  movel([0.147187, -1.292502, -2.622642, -0.797245, 1.570796, 1.717984],accel_mss,speed_ms,0,blend_radius_m)
  movel([0.147550, -1.292939, -2.622384, -0.797065, 1.570796, 1.718347],accel_mss,speed_ms,0,blend_radius_m)
  movel([0.147774, -1.294240, -2.621617, -0.796531, 1.570796, 1.718570],accel_mss,speed_ms,0,blend_radius_m)
  movel([0.147672, -1.296185, -2.620466, -0.795737, 1.570796, 1.718469],accel_mss,speed_ms,0,blend_radius_m)
  movel([0.147381, -1.298185, -2.619278, -0.794926, 1.570796, 1.718178],accel_mss,speed_ms,0,blend_radius_m)
  movel([0.149143, -1.296279, -2.620411, -0.795699, 1.570796, 1.719939],accel_mss,speed_ms,0,blend_radius_m)
  movel([0.151055, -1.294467, -2.621483, -0.796439, 1.570796, 1.721852],accel_mss,speed_ms,0,blend_radius_m)
  movel([0.153085, -1.292767, -2.622486, -0.797136, 1.570796, 1.723882],accel_mss,speed_ms,0,blend_radius_m)
  movel([0.155193, -1.291198, -2.623408, -0.797783, 1.570796, 1.725989],accel_mss,speed_ms,0,blend_radius_m)
  movel([0.159402, -1.288061, -2.625242, -0.799086, 1.570796, 1.730199],accel_mss,speed_ms,0,blend_radius_m)
  movel([0.160619, -1.287255, -2.625711, -0.799423, 1.570796, 1.731416],accel_mss,speed_ms,0,blend_radius_m)
  movel([0.161780, -1.286599, -2.626092, -0.799698, 1.570796, 1.732576],accel_mss,speed_ms,0,blend_radius_m)
  movel([0.162826, -1.286172, -2.626340, -0.799877, 1.570796, 1.733623],accel_mss,speed_ms,0,blend_radius_m)
  movel([0.163696, -1.286049, -2.626411, -0.799928, 1.570796, 1.734492],accel_mss,speed_ms,0,blend_radius_m)
  movel([0.164332, -1.286333, -2.626247, -0.799809, 1.570796, 1.735128],accel_mss,speed_ms,0,blend_radius_m)
  movel([0.164662, -1.286984, -2.625868, -0.799536, 1.570796, 1.735459],accel_mss,speed_ms,0,blend_radius_m)
  movel([0.164729, -1.287902, -2.625335, -0.799153, 1.570796, 1.735526],accel_mss,speed_ms,0,blend_radius_m)
  movel([0.164568, -1.288980, -2.624706, -0.798703, 1.570796, 1.735364],accel_mss,speed_ms,0,blend_radius_m)
  movel([0.164219, -1.290117, -2.624041, -0.798231, 1.570796, 1.735015],accel_mss,speed_ms,0,blend_radius_m)
  movel([0.163722, -1.291209, -2.623401, -0.797779, 1.570796, 1.734518],accel_mss,speed_ms,0,blend_radius_m)
  movel([0.163113, -1.292155, -2.622846, -0.797388, 1.570796, 1.733910],accel_mss,speed_ms,0,blend_radius_m)
  movel([0.162431, -1.292853, -2.622435, -0.797101, 1.570796, 1.733227],accel_mss,speed_ms,0,blend_radius_m)
  movel([0.166229, -1.290188, -2.624000, -0.798201, 1.570796, 1.737025],accel_mss,speed_ms,0,blend_radius_m)
  movel([0.168191, -1.288999, -2.624694, -0.798695, 1.570796, 1.738988],accel_mss,speed_ms,0,blend_radius_m)
  movel([0.170182, -1.287929, -2.625319, -0.799141, 1.570796, 1.740979],accel_mss,speed_ms,0,blend_radius_m)
  movel([0.172188, -1.286991, -2.625865, -0.799534, 1.570796, 1.742984],accel_mss,speed_ms,0,blend_radius_m)
  movel([0.174199, -1.286202, -2.626323, -0.799864, 1.570796, 1.744995],accel_mss,speed_ms,0,blend_radius_m)
  movel([0.176204, -1.285580, -2.626683, -0.800126, 1.570796, 1.747000],accel_mss,speed_ms,0,blend_radius_m)
  movel([0.178191, -1.285136, -2.626940, -0.800312, 1.570796, 1.748987],accel_mss,speed_ms,0,blend_radius_m)
  movel([0.179463, -1.285131, -2.626943, -0.800314, 1.570796, 1.750259],accel_mss,speed_ms,0,blend_radius_m)
  movel([0.180721, -1.285520, -2.626718, -0.800151, 1.570796, 1.751518],accel_mss,speed_ms,0,blend_radius_m)
  movel([0.181223, -1.285864, -2.626519, -0.800006, 1.570796, 1.752019],accel_mss,speed_ms,0,blend_radius_m)
  movel([0.181576, -1.286307, -2.626262, -0.799820, 1.570796, 1.752372],accel_mss,speed_ms,0,blend_radius_m)
  movel([0.181734, -1.286851, -2.625946, -0.799592, 1.570796, 1.752530],accel_mss,speed_ms,0,blend_radius_m)
  movel([0.181645, -1.287496, -2.625571, -0.799322, 1.570796, 1.752441],accel_mss,speed_ms,0,blend_radius_m)
  movel([0.181300, -1.288146, -2.625192, -0.799051, 1.570796, 1.752096],accel_mss,speed_ms,0,blend_radius_m)
  movel([0.180775, -1.288760, -2.624834, -0.798795, 1.570796, 1.751571],accel_mss,speed_ms,0,blend_radius_m)
  movel([0.179372, -1.289953, -2.624137, -0.798299, 1.570796, 1.750168],accel_mss,speed_ms,0,blend_radius_m)
  movel([0.177819, -1.290875, -2.623597, -0.797917, 1.570796, 1.748615],accel_mss,speed_ms,0,blend_radius_m)
  movel([0.176195, -1.291571, -2.623189, -0.797629, 1.570796, 1.746991],accel_mss,speed_ms,0,blend_radius_m)
  movel([0.174578, -1.292087, -2.622886, -0.797416, 1.570796, 1.745374],accel_mss,speed_ms,0,blend_radius_m)
  movel([0.176378, -1.292531, -2.622625, -0.797233, 1.570796, 1.747174],accel_mss,speed_ms,0,blend_radius_m)
  movel([0.178306, -1.292768, -2.622485, -0.797136, 1.570796, 1.749103],accel_mss,speed_ms,0,blend_radius_m)
  movel([0.180340, -1.292800, -2.622467, -0.797123, 1.570796, 1.751137],accel_mss,speed_ms,0,blend_radius_m)
  movel([0.182461, -1.292627, -2.622568, -0.797194, 1.570796, 1.753257],accel_mss,speed_ms,0,blend_radius_m)
  movel([0.184182, -1.292297, -2.622762, -0.797330, 1.570796, 1.754979],accel_mss,speed_ms,0,blend_radius_m)
  movel([0.187621, -1.291362, -2.623311, -0.797715, 1.570796, 1.758417],accel_mss,speed_ms,0,blend_radius_m)
  movel([0.189347, -1.291019, -2.623513, -0.797857, 1.570796, 1.760143],accel_mss,speed_ms,0,blend_radius_m)
  movel([0.191271, -1.290783, -2.623651, -0.797955, 1.570796, 1.762067],accel_mss,speed_ms,0,blend_radius_m)
  movel([0.194455, -1.290577, -2.623772, -0.798040, 1.570796, 1.765251],accel_mss,speed_ms,0,blend_radius_m)
  movel([0.195937, -1.290628, -2.623742, -0.798019, 1.570796, 1.766733],accel_mss,speed_ms,0,blend_radius_m)
  movel([0.197036, -1.290857, -2.623608, -0.797924, 1.570796, 1.767833],accel_mss,speed_ms,0,blend_radius_m)
  movel([0.197371, -1.291056, -2.623491, -0.797842, 1.570796, 1.768167],accel_mss,speed_ms,0,blend_radius_m)
  movel([0.197521, -1.291320, -2.623336, -0.797733, 1.570796, 1.768317],accel_mss,speed_ms,0,blend_radius_m)
  movel([0.197462, -1.291654, -2.623140, -0.797595, 1.570796, 1.768258],accel_mss,speed_ms,0,blend_radius_m)
  movel([0.197162, -1.292065, -2.622898, -0.797425, 1.570796, 1.767958],accel_mss,speed_ms,0,blend_radius_m)
  movel([0.196189, -1.292919, -2.622396, -0.797073, 1.570796, 1.766986],accel_mss,speed_ms,0,blend_radius_m)
  movel([0.195007, -1.293687, -2.621944, -0.796758, 1.570796, 1.765803],accel_mss,speed_ms,0,blend_radius_m)
  movel([0.193677, -1.294378, -2.621536, -0.796475, 1.570796, 1.764473],accel_mss,speed_ms,0,blend_radius_m)
  movel([0.192268, -1.294993, -2.621172, -0.796224, 1.570796, 1.763065],accel_mss,speed_ms,0,blend_radius_m)
  movel([0.189469, -1.296012, -2.620569, -0.795808, 1.570796, 1.760265],accel_mss,speed_ms,0,blend_radius_m)
  movel([0.187130, -1.296774, -2.620117, -0.795498, 1.570796, 1.757926],accel_mss,speed_ms,0,blend_radius_m)
  movel([0.188093, -1.297277, -2.619818, -0.795294, 1.570796, 1.758889],accel_mss,speed_ms,0,blend_radius_m)
  movel([0.189142, -1.297667, -2.619586, -0.795136, 1.570796, 1.759938],accel_mss,speed_ms,0,blend_radius_m)
  movel([0.191445, -1.298162, -2.619291, -0.794935, 1.570796, 1.762241],accel_mss,speed_ms,0,blend_radius_m)
  movel([0.193943, -1.298359, -2.619175, -0.794856, 1.570796, 1.764739],accel_mss,speed_ms,0,blend_radius_m)
  movel([0.196543, -1.298358, -2.619175, -0.794856, 1.570796, 1.767339],accel_mss,speed_ms,0,blend_radius_m)
  movel([0.198733, -1.298215, -2.619260, -0.794914, 1.570796, 1.769529],accel_mss,speed_ms,0,blend_radius_m)
  movel([0.205405, -1.297512, -2.619678, -0.795198, 1.570796, 1.776202],accel_mss,speed_ms,0,blend_radius_m)
  movel([0.206582, -1.297609, -2.619621, -0.795159, 1.570796, 1.777379],accel_mss,speed_ms,0,blend_radius_m)
  movel([0.207429, -1.297998, -2.619389, -0.795002, 1.570796, 1.778225],accel_mss,speed_ms,0,blend_radius_m)
  movel([0.207554, -1.298296, -2.619212, -0.794881, 1.570796, 1.778350],accel_mss,speed_ms,0,blend_radius_m)
  movel([0.207384, -1.298662, -2.618994, -0.794733, 1.570796, 1.778180],accel_mss,speed_ms,0,blend_radius_m)
  movel([0.206850, -1.299092, -2.618737, -0.794560, 1.570796, 1.777646],accel_mss,speed_ms,0,blend_radius_m)
  movel([0.205881, -1.299582, -2.618444, -0.794362, 1.570796, 1.776677],accel_mss,speed_ms,0,blend_radius_m)
  movel([0.204309, -1.300170, -2.618093, -0.794126, 1.570796, 1.775105],accel_mss,speed_ms,0,blend_radius_m)
  movel([0.202535, -1.300655, -2.617803, -0.793931, 1.570796, 1.773331],accel_mss,speed_ms,0,blend_radius_m)
  movel([0.200836, -1.300909, -2.617651, -0.793829, 1.570796, 1.771632],accel_mss,speed_ms,0,blend_radius_m)
  movel([0.200100, -1.300910, -2.617650, -0.793829, 1.570796, 1.770896],accel_mss,speed_ms,0,blend_radius_m)
  movel([0.199490, -1.300801, -2.617716, -0.793873, 1.570796, 1.770286],accel_mss,speed_ms,0,blend_radius_m)
  movel([0.201611, -1.302312, -2.616809, -0.793268, 1.570796, 1.772407],accel_mss,speed_ms,0,blend_radius_m)
  movel([0.203973, -1.303547, -2.616066, -0.792776, 1.570796, 1.774769],accel_mss,speed_ms,0,blend_radius_m)
  movel([0.206525, -1.304557, -2.615457, -0.792375, 1.570796, 1.777321],accel_mss,speed_ms,0,blend_radius_m)
  movel([0.209220, -1.305396, -2.614950, -0.792043, 1.570796, 1.780016],accel_mss,speed_ms,0,blend_radius_m)
  movel([0.214839, -1.306755, -2.614126, -0.791507, 1.570796, 1.785635],accel_mss,speed_ms,0,blend_radius_m)
  movel([0.220430, -1.308023, -2.613356, -0.791010, 1.570796, 1.791226],accel_mss,speed_ms,0,blend_radius_m)
  movel([0.221316, -1.308412, -2.613120, -0.790858, 1.570796, 1.792112],accel_mss,speed_ms,0,blend_radius_m)
  movel([0.221557, -1.308760, -2.612908, -0.790722, 1.570796, 1.792354],accel_mss,speed_ms,0,blend_radius_m)
  movel([0.221539, -1.309244, -2.612612, -0.790532, 1.570796, 1.792335],accel_mss,speed_ms,0,blend_radius_m)
  movel([0.221247, -1.309765, -2.612295, -0.790329, 1.570796, 1.792044],accel_mss,speed_ms,0,blend_radius_m)
  movel([0.220033, -1.310912, -2.611593, -0.789884, 1.570796, 1.790829],accel_mss,speed_ms,0,blend_radius_m)
  movel([0.219216, -1.311486, -2.611242, -0.789661, 1.570796, 1.790013],accel_mss,speed_ms,0,blend_radius_m)
  movel([0.217461, -1.312385, -2.610691, -0.789314, 1.570796, 1.788257],accel_mss,speed_ms,0,blend_radius_m)
  movel([0.215610, -1.312982, -2.610324, -0.789083, 1.570796, 1.786407],accel_mss,speed_ms,0,blend_radius_m)
  movel([0.213729, -1.313322, -2.610115, -0.788953, 1.570796, 1.784525],accel_mss,speed_ms,0,blend_radius_m)
  movel([0.211888, -1.313440, -2.610042, -0.788907, 1.570796, 1.782685],accel_mss,speed_ms,0,blend_radius_m)
  movel([0.210157, -1.313379, -2.610079, -0.788930, 1.570796, 1.780953],accel_mss,speed_ms,0,blend_radius_m)
  movel([0.208604, -1.313175, -2.610205, -0.789009, 1.570796, 1.779400],accel_mss,speed_ms,0,blend_radius_m)
  movel([0.207302, -1.312863, -2.610397, -0.789129, 1.570796, 1.778098],accel_mss,speed_ms,0,blend_radius_m)
  movel([0.207188, -1.313311, -2.610121, -0.788957, 1.570796, 1.777984],accel_mss,speed_ms,0,blend_radius_m)
  movel([0.207346, -1.313680, -2.609894, -0.788815, 1.570796, 1.778142],accel_mss,speed_ms,0,blend_radius_m)
  movel([0.207939, -1.314359, -2.609476, -0.788554, 1.570796, 1.778735],accel_mss,speed_ms,0,blend_radius_m)
  movel([0.208657, -1.314923, -2.609128, -0.788338, 1.570796, 1.779454],accel_mss,speed_ms,0,blend_radius_m)
  movel([0.210309, -1.315835, -2.608564, -0.787990, 1.570796, 1.781105],accel_mss,speed_ms,0,blend_radius_m)
  movel([0.213305, -1.317223, -2.607704, -0.787461, 1.570796, 1.784102],accel_mss,speed_ms,0,blend_radius_m)
  movel([0.216384, -1.318478, -2.606925, -0.786986, 1.570796, 1.787181],accel_mss,speed_ms,0,blend_radius_m)
  movel([0.222772, -1.320657, -2.605566, -0.786166, 1.570796, 1.793568],accel_mss,speed_ms,0,blend_radius_m)
  movel([0.224533, -1.321298, -2.605165, -0.785925, 1.570796, 1.795329],accel_mss,speed_ms,0,blend_radius_m)
  movel([0.225622, -1.321824, -2.604836, -0.785729, 1.570796, 1.796418],accel_mss,speed_ms,0,blend_radius_m)
  movel([0.226633, -1.322477, -2.604427, -0.785485, 1.570796, 1.797429],accel_mss,speed_ms,0,blend_radius_m)
  movel([0.227396, -1.323251, -2.603940, -0.785197, 1.570796, 1.798192],accel_mss,speed_ms,0,blend_radius_m)
  movel([0.227749, -1.324134, -2.603385, -0.784870, 1.570796, 1.798546],accel_mss,speed_ms,0,blend_radius_m)
  movel([0.227725, -1.324612, -2.603084, -0.784693, 1.570796, 1.798521],accel_mss,speed_ms,0,blend_radius_m)
  movel([0.227538, -1.325115, -2.602767, -0.784507, 1.570796, 1.798334],accel_mss,speed_ms,0,blend_radius_m)
  movel([0.227164, -1.325643, -2.602434, -0.784312, 1.570796, 1.797961],accel_mss,speed_ms,0,blend_radius_m)
  movel([0.226591, -1.326191, -2.602087, -0.784110, 1.570796, 1.797387],accel_mss,speed_ms,0,blend_radius_m)
  movel([0.225837, -1.326540, -2.601867, -0.783982, 1.570796, 1.796634],accel_mss,speed_ms,0,blend_radius_m)
  movel([0.224871, -1.326699, -2.601766, -0.783924, 1.570796, 1.795668],accel_mss,speed_ms,0,blend_radius_m)
  movel([0.219802, -1.326944, -2.601611, -0.783834, 1.570796, 1.790598],accel_mss,speed_ms,0,blend_radius_m)
  movel([0.218145, -1.326787, -2.601710, -0.783892, 1.570796, 1.788941],accel_mss,speed_ms,0,blend_radius_m)
  movel([0.217459, -1.326589, -2.601836, -0.783964, 1.570796, 1.788255],accel_mss,speed_ms,0,blend_radius_m)
  movel([0.216923, -1.326283, -2.602029, -0.784077, 1.570796, 1.787719],accel_mss,speed_ms,0,blend_radius_m)
  movel([0.218941, -1.328596, -2.600563, -0.783230, 1.570796, 1.789737],accel_mss,speed_ms,0,blend_radius_m)
  movel([0.221308, -1.330580, -2.599299, -0.782510, 1.570796, 1.792105],accel_mss,speed_ms,0,blend_radius_m)
  movel([0.223948, -1.332287, -2.598208, -0.781894, 1.570796, 1.794744],accel_mss,speed_ms,0,blend_radius_m)
  movel([0.226784, -1.333763, -2.597261, -0.781365, 1.570796, 1.797581],accel_mss,speed_ms,0,blend_radius_m)
  movel([0.229318, -1.334606, -2.596719, -0.781064, 1.570796, 1.800115],accel_mss,speed_ms,0,blend_radius_m)
  movel([0.232932, -1.335887, -2.595893, -0.780608, 1.570796, 1.803728],accel_mss,speed_ms,0,blend_radius_m)
  movel([0.234525, -1.336695, -2.595372, -0.780322, 1.570796, 1.805322],accel_mss,speed_ms,0,blend_radius_m)
  movel([0.235653, -1.337610, -2.594780, -0.780000, 1.570796, 1.806450],accel_mss,speed_ms,0,blend_radius_m)
  movel([0.235966, -1.338106, -2.594458, -0.779825, 1.570796, 1.806763],accel_mss,speed_ms,0,blend_radius_m)
  movel([0.236070, -1.338627, -2.594120, -0.779642, 1.570796, 1.806867],accel_mss,speed_ms,0,blend_radius_m)
  movel([0.235936, -1.339175, -2.593764, -0.779450, 1.570796, 1.806733],accel_mss,speed_ms,0,blend_radius_m)
  movel([0.235538, -1.339746, -2.593393, -0.779250, 1.570796, 1.806335],accel_mss,speed_ms,0,blend_radius_m)
  movel([0.234996, -1.340245, -2.593068, -0.779076, 1.570796, 1.805793],accel_mss,speed_ms,0,blend_radius_m)
  movel([0.234397, -1.340669, -2.592792, -0.778928, 1.570796, 1.805193],accel_mss,speed_ms,0,blend_radius_m)
  movel([0.233113, -1.341353, -2.592346, -0.778690, 1.570796, 1.803910],accel_mss,speed_ms,0,blend_radius_m)
  movel([0.231720, -1.341950, -2.591956, -0.778483, 1.570796, 1.802517],accel_mss,speed_ms,0,blend_radius_m)
  movel([0.228948, -1.342826, -2.591382, -0.778180, 1.570796, 1.799744],accel_mss,speed_ms,0,blend_radius_m)
  movel([0.227584, -1.343104, -2.591201, -0.778085, 1.570796, 1.798381],accel_mss,speed_ms,0,blend_radius_m)
  movel([0.229786, -1.344148, -2.590516, -0.777725, 1.570796, 1.800582],accel_mss,speed_ms,0,blend_radius_m)
  movel([0.232093, -1.345031, -2.589935, -0.777422, 1.570796, 1.802889],accel_mss,speed_ms,0,blend_radius_m)
  movel([0.234492, -1.345775, -2.589446, -0.777168, 1.570796, 1.805289],accel_mss,speed_ms,0,blend_radius_m)
  movel([0.236975, -1.346392, -2.589039, -0.776958, 1.570796, 1.807771],accel_mss,speed_ms,0,blend_radius_m)
  movel([0.242140, -1.347324, -2.588424, -0.776642, 1.570796, 1.812936],accel_mss,speed_ms,0,blend_radius_m)
  movel([0.247502, -1.347956, -2.588005, -0.776427, 1.570796, 1.818298],accel_mss,speed_ms,0,blend_radius_m)
  movel([0.248879, -1.348279, -2.587792, -0.776318, 1.570796, 1.819675],accel_mss,speed_ms,0,blend_radius_m)
  movel([0.249326, -1.348656, -2.587542, -0.776191, 1.570796, 1.820123],accel_mss,speed_ms,0,blend_radius_m)
  movel([0.249438, -1.349252, -2.587147, -0.775991, 1.570796, 1.820234],accel_mss,speed_ms,0,blend_radius_m)
  movel([0.249300, -1.349711, -2.586842, -0.775836, 1.570796, 1.820097],accel_mss,speed_ms,0,blend_radius_m)
  movel([0.249032, -1.350158, -2.586545, -0.775686, 1.570796, 1.819828],accel_mss,speed_ms,0,blend_radius_m)
  movel([0.248159, -1.351020, -2.585971, -0.775398, 1.570796, 1.818956],accel_mss,speed_ms,0,blend_radius_m)
  movel([0.246957, -1.351813, -2.585442, -0.775133, 1.570796, 1.817753],accel_mss,speed_ms,0,blend_radius_m)
  movel([0.245556, -1.352524, -2.584968, -0.774897, 1.570796, 1.816352],accel_mss,speed_ms,0,blend_radius_m)
  movel([0.242697, -1.353616, -2.584238, -0.774536, 1.570796, 1.813494],accel_mss,speed_ms,0,blend_radius_m)
  movel([0.240653, -1.354136, -2.583889, -0.774364, 1.570796, 1.811449],accel_mss,speed_ms,0,blend_radius_m)
  movel([0.241713, -1.354387, -2.583721, -0.774281, 1.570796, 1.812509],accel_mss,speed_ms,0,blend_radius_m)
  movel([0.242833, -1.354526, -2.583627, -0.774235, 1.570796, 1.813629],accel_mss,speed_ms,0,blend_radius_m)
  movel([0.245219, -1.354502, -2.583643, -0.774243, 1.570796, 1.816016],accel_mss,speed_ms,0,blend_radius_m)
  movel([0.247757, -1.354097, -2.583915, -0.774377, 1.570796, 1.818553],accel_mss,speed_ms,0,blend_radius_m)
  movel([0.250387, -1.353354, -2.584413, -0.774622, 1.570796, 1.821184],accel_mss,speed_ms,0,blend_radius_m)
  movel([0.253059, -1.352300, -2.585117, -0.774971, 1.570796, 1.823855],accel_mss,speed_ms,0,blend_radius_m)
  movel([0.255714, -1.350980, -2.585997, -0.775411, 1.570796, 1.826510],accel_mss,speed_ms,0,blend_radius_m)
  movel([0.258298, -1.349422, -2.587033, -0.775933, 1.570796, 1.829094],accel_mss,speed_ms,0,blend_radius_m)
  movel([0.260755, -1.347666, -2.588197, -0.776526, 1.570796, 1.831551],accel_mss,speed_ms,0,blend_radius_m)
  movel([0.261839, -1.346878, -2.588718, -0.776793, 1.570796, 1.832635],accel_mss,speed_ms,0,blend_radius_m)
  movel([0.262400, -1.346588, -2.588910, -0.776891, 1.570796, 1.833196],accel_mss,speed_ms,0,blend_radius_m)
  movel([0.262957, -1.346439, -2.589008, -0.776942, 1.570796, 1.833753],accel_mss,speed_ms,0,blend_radius_m)
  movel([0.263495, -1.346496, -2.588970, -0.776923, 1.570796, 1.834292],accel_mss,speed_ms,0,blend_radius_m)
  movel([0.263919, -1.346727, -2.588818, -0.776844, 1.570796, 1.834715],accel_mss,speed_ms,0,blend_radius_m)
  movel([0.264319, -1.347325, -2.588423, -0.776641, 1.570796, 1.835115],accel_mss,speed_ms,0,blend_radius_m)
  movel([0.264431, -1.348166, -2.587866, -0.776356, 1.570796, 1.835227],accel_mss,speed_ms,0,blend_radius_m)
  movel([0.264312, -1.349180, -2.587194, -0.776015, 1.570796, 1.835108],accel_mss,speed_ms,0,blend_radius_m)
  movel([0.264015, -1.350302, -2.586449, -0.775638, 1.570796, 1.834811],accel_mss,speed_ms,0,blend_radius_m)
  movel([0.263105, -1.352585, -2.584927, -0.774877, 1.570796, 1.833901],accel_mss,speed_ms,0,blend_radius_m)
  movel([0.262138, -1.354477, -2.583660, -0.774252, 1.570796, 1.832934],accel_mss,speed_ms,0,blend_radius_m)
  movel([0.264294, -1.352626, -2.584900, -0.774863, 1.570796, 1.835090],accel_mss,speed_ms,0,blend_radius_m)
  movel([0.266279, -1.350629, -2.586232, -0.775529, 1.570796, 1.837075],accel_mss,speed_ms,0,blend_radius_m)
  movel([0.268078, -1.348508, -2.587640, -0.776241, 1.570796, 1.838874],accel_mss,speed_ms,0,blend_radius_m)
  movel([0.269679, -1.346299, -2.589100, -0.776990, 1.570796, 1.840475],accel_mss,speed_ms,0,blend_radius_m)
  movel([0.271060, -1.344027, -2.590595, -0.777767, 1.570796, 1.841856],accel_mss,speed_ms,0,blend_radius_m)
  movel([0.272215, -1.341720, -2.592106, -0.778563, 1.570796, 1.843011],accel_mss,speed_ms,0,blend_radius_m)
  movel([0.273119, -1.339412, -2.593610, -0.779367, 1.570796, 1.843916],accel_mss,speed_ms,0,blend_radius_m)
  movel([0.273761, -1.337131, -2.595089, -0.780168, 1.570796, 1.844557],accel_mss,speed_ms,0,blend_radius_m)
  movel([0.274224, -1.334033, -2.597088, -0.781268, 1.570796, 1.845020],accel_mss,speed_ms,0,blend_radius_m)
  movel([0.274591, -1.332385, -2.598145, -0.781859, 1.570796, 1.845387],accel_mss,speed_ms,0,blend_radius_m)
  movel([0.274879, -1.331604, -2.598645, -0.782140, 1.570796, 1.845675],accel_mss,speed_ms,0,blend_radius_m)
  movel([0.275260, -1.330877, -2.599109, -0.782402, 1.570796, 1.846056],accel_mss,speed_ms,0,blend_radius_m)
  movel([0.276072, -1.329798, -2.599798, -0.782793, 1.570796, 1.846868],accel_mss,speed_ms,0,blend_radius_m)
  movel([0.276761, -1.329255, -2.600144, -0.782990, 1.570796, 1.847557],accel_mss,speed_ms,0,blend_radius_m)
  movel([0.277351, -1.329134, -2.600221, -0.783034, 1.570796, 1.848147],accel_mss,speed_ms,0,blend_radius_m)
  movel([0.277863, -1.329315, -2.600105, -0.782968, 1.570796, 1.848659],accel_mss,speed_ms,0,blend_radius_m)
  movel([0.279119, -1.330501, -2.599350, -0.782538, 1.570796, 1.849916],accel_mss,speed_ms,0,blend_radius_m)
  movel([0.279515, -1.330717, -2.599212, -0.782460, 1.570796, 1.850311],accel_mss,speed_ms,0,blend_radius_m)
  movel([0.280667, -1.329098, -2.600244, -0.783047, 1.570796, 1.851463],accel_mss,speed_ms,0,blend_radius_m)
  movel([0.281683, -1.327421, -2.601309, -0.783659, 1.570796, 1.852479],accel_mss,speed_ms,0,blend_radius_m)
  movel([0.282568, -1.325699, -2.602399, -0.784292, 1.570796, 1.853364],accel_mss,speed_ms,0,blend_radius_m)
  movel([0.283329, -1.323939, -2.603508, -0.784942, 1.570796, 1.854125],accel_mss,speed_ms,0,blend_radius_m)
  movel([0.283966, -1.322154, -2.604629, -0.785606, 1.570796, 1.854762],accel_mss,speed_ms,0,blend_radius_m)
  movel([0.284486, -1.320354, -2.605755, -0.786279, 1.570796, 1.855282],accel_mss,speed_ms,0,blend_radius_m)
  movel([0.285202, -1.316750, -2.607998, -0.787641, 1.570796, 1.855998],accel_mss,speed_ms,0,blend_radius_m)
  movel([0.285512, -1.313217, -2.610179, -0.788993, 1.570796, 1.856308],accel_mss,speed_ms,0,blend_radius_m)
  movel([0.285464, -1.309843, -2.612247, -0.790299, 1.570796, 1.856260],accel_mss,speed_ms,0,blend_radius_m)
  movel([0.285091, -1.306721, -2.614147, -0.791521, 1.570796, 1.855888],accel_mss,speed_ms,0,blend_radius_m)
  movel([0.284446, -1.303940, -2.615829, -0.792620, 1.570796, 1.855243],accel_mss,speed_ms,0,blend_radius_m)
  speed_ms = 0.005
  movel([0.284446, -1.294903, -2.611476, -0.806009, 1.570796, 1.855243],accel_mss,speed_ms,0,blend_radius_m)
  speed_ms = 0.040
  movel([0.269748, -1.298612, -2.609260, -0.804517, 1.570796, 1.840544],accel_mss,speed_ms,0,blend_radius_m)
  speed_ms = 0.005
  movel([0.269748, -1.307628, -2.613596, -0.791164, 1.570796, 1.840544],accel_mss,speed_ms,0,blend_radius_m)
  speed_ms = 0.025
  movel([0.268699, -1.306702, -2.614159, -0.791528, 1.570796, 1.839496],accel_mss,speed_ms,0,blend_radius_m)
  movel([0.267398, -1.306097, -2.614525, -0.791766, 1.570796, 1.838194],accel_mss,speed_ms,0,blend_radius_m)
  movel([0.265889, -1.305774, -2.614721, -0.791894, 1.570796, 1.836685],accel_mss,speed_ms,0,blend_radius_m)
  movel([0.264223, -1.305688, -2.614773, -0.791928, 1.570796, 1.835020],accel_mss,speed_ms,0,blend_radius_m)
  movel([0.262449, -1.305799, -2.614706, -0.791884, 1.570796, 1.833245],accel_mss,speed_ms,0,blend_radius_m)
  movel([0.260612, -1.306063, -2.614546, -0.791780, 1.570796, 1.831408],accel_mss,speed_ms,0,blend_radius_m)
  movel([0.256944, -1.306876, -2.614053, -0.791460, 1.570796, 1.827740],accel_mss,speed_ms,0,blend_radius_m)
  speed_ms = 0.005
  movel([0.256944, -1.297855, -2.609714, -0.804820, 1.570796, 1.827740],accel_mss,speed_ms,0,blend_radius_m)
  speed_ms = 0.040
  movel([0.261759, -1.296351, -2.610614, -0.805425, 1.570796, 1.832555],accel_mss,speed_ms,0,blend_radius_m)
  speed_ms = 0.005
  movel([0.261759, -1.305379, -2.614960, -0.792050, 1.570796, 1.832555],accel_mss,speed_ms,0,blend_radius_m)
  speed_ms = 0.025
  movel([0.262808, -1.303409, -2.616149, -0.792831, 1.570796, 1.833605],accel_mss,speed_ms,0,blend_radius_m)
  movel([0.263652, -1.301488, -2.617304, -0.793597, 1.570796, 1.834449],accel_mss,speed_ms,0,blend_radius_m)
  movel([0.264295, -1.299615, -2.618425, -0.794349, 1.570796, 1.835092],accel_mss,speed_ms,0,blend_radius_m)
  movel([0.264748, -1.297784, -2.619517, -0.795088, 1.570796, 1.835544],accel_mss,speed_ms,0,blend_radius_m)
  movel([0.265022, -1.295992, -2.620581, -0.795816, 1.570796, 1.835819],accel_mss,speed_ms,0,blend_radius_m)
  movel([0.265127, -1.294235, -2.621620, -0.796534, 1.570796, 1.835923],accel_mss,speed_ms,0,blend_radius_m)
  movel([0.265071, -1.292510, -2.622637, -0.797242, 1.570796, 1.835868],accel_mss,speed_ms,0,blend_radius_m)
  movel([0.264867, -1.290813, -2.623634, -0.797943, 1.570796, 1.835663],accel_mss,speed_ms,0,blend_radius_m)
  movel([0.263809, -1.286044, -2.626414, -0.799931, 1.570796, 1.834606],accel_mss,speed_ms,0,blend_radius_m)
  movel([0.263405, -1.283705, -2.627768, -0.800916, 1.570796, 1.834201],accel_mss,speed_ms,0,blend_radius_m)
  movel([0.263315, -1.280988, -2.629331, -0.802070, 1.570796, 1.834111],accel_mss,speed_ms,0,blend_radius_m)
  movel([0.263585, -1.277432, -2.631364, -0.803594, 1.570796, 1.834381],accel_mss,speed_ms,0,blend_radius_m)
  movel([0.264171, -1.273757, -2.633447, -0.805185, 1.570796, 1.834967],accel_mss,speed_ms,0,blend_radius_m)
  movel([0.265168, -1.269976, -2.635574, -0.806840, 1.570796, 1.835964],accel_mss,speed_ms,0,blend_radius_m)
  movel([0.265850, -1.268048, -2.636651, -0.807690, 1.570796, 1.836646],accel_mss,speed_ms,0,blend_radius_m)
  movel([0.266671, -1.266100, -2.637735, -0.808554, 1.570796, 1.837468],accel_mss,speed_ms,0,blend_radius_m)
  movel([0.268233, -1.263113, -2.639388, -0.809888, 1.570796, 1.839029],accel_mss,speed_ms,0,blend_radius_m)
  movel([0.270105, -1.260274, -2.640949, -0.811166, 1.570796, 1.840901],accel_mss,speed_ms,0,blend_radius_m)
  movel([0.272263, -1.257600, -2.642411, -0.812379, 1.570796, 1.843059],accel_mss,speed_ms,0,blend_radius_m)
  movel([0.274682, -1.255112, -2.643763, -0.813514, 1.570796, 1.845478],accel_mss,speed_ms,0,blend_radius_m)
  movel([0.277330, -1.252836, -2.644993, -0.814560, 1.570796, 1.848127],accel_mss,speed_ms,0,blend_radius_m)
  movel([0.280184, -1.250792, -2.646092, -0.815504, 1.570796, 1.850980],accel_mss,speed_ms,0,blend_radius_m)
  movel([0.283216, -1.249001, -2.647052, -0.816336, 1.570796, 1.854012],accel_mss,speed_ms,0,blend_radius_m)
  movel([0.286392, -1.247489, -2.647859, -0.817041, 1.570796, 1.857188],accel_mss,speed_ms,0,blend_radius_m)
  movel([0.288816, -1.246569, -2.648348, -0.817471, 1.570796, 1.859612],accel_mss,speed_ms,0,blend_radius_m)
  movel([0.291238, -1.245851, -2.648730, -0.817808, 1.570796, 1.862034],accel_mss,speed_ms,0,blend_radius_m)
  movel([0.293635, -1.245335, -2.649004, -0.818050, 1.570796, 1.864431],accel_mss,speed_ms,0,blend_radius_m)
  movel([0.295991, -1.245016, -2.649173, -0.818200, 1.570796, 1.866788],accel_mss,speed_ms,0,blend_radius_m)
  movel([0.298283, -1.244900, -2.649234, -0.818255, 1.570796, 1.869079],accel_mss,speed_ms,0,blend_radius_m)
  movel([0.300490, -1.244983, -2.649190, -0.818216, 1.570796, 1.871287],accel_mss,speed_ms,0,blend_radius_m)
  movel([0.302592, -1.245263, -2.649042, -0.818084, 1.570796, 1.873389],accel_mss,speed_ms,0,blend_radius_m)
  movel([0.304570, -1.245741, -2.648788, -0.817860, 1.570796, 1.875366],accel_mss,speed_ms,0,blend_radius_m)
  movel([0.306400, -1.246413, -2.648431, -0.817544, 1.570796, 1.877196],accel_mss,speed_ms,0,blend_radius_m)
  movel([0.308069, -1.247277, -2.647972, -0.817140, 1.570796, 1.878865],accel_mss,speed_ms,0,blend_radius_m)
  movel([0.309554, -1.248331, -2.647410, -0.816648, 1.570796, 1.880350],accel_mss,speed_ms,0,blend_radius_m)
  movel([0.310838, -1.249571, -2.646747, -0.816071, 1.570796, 1.881635],accel_mss,speed_ms,0,blend_radius_m)
  movel([0.311904, -1.250993, -2.645984, -0.815411, 1.570796, 1.882700],accel_mss,speed_ms,0,blend_radius_m)
  movel([0.312728, -1.252597, -2.645122, -0.814670, 1.570796, 1.883525],accel_mss,speed_ms,0,blend_radius_m)
  movel([0.313299, -1.254374, -2.644162, -0.813853, 1.570796, 1.884095],accel_mss,speed_ms,0,blend_radius_m)
  movel([0.313596, -1.256325, -2.643104, -0.812960, 1.570796, 1.884393],accel_mss,speed_ms,0,blend_radius_m)
  movel([0.313652, -1.259020, -2.641636, -0.811734, 1.570796, 1.884448],accel_mss,speed_ms,0,blend_radius_m)
  movel([0.313460, -1.261807, -2.640107, -0.810475, 1.570796, 1.884256],accel_mss,speed_ms,0,blend_radius_m)
  movel([0.313070, -1.264658, -2.638534, -0.809197, 1.570796, 1.883867],accel_mss,speed_ms,0,blend_radius_m)
  movel([0.312543, -1.267539, -2.636935, -0.807916, 1.570796, 1.883339],accel_mss,speed_ms,0,blend_radius_m)
  movel([0.311121, -1.273822, -2.633411, -0.805157, 1.570796, 1.881917],accel_mss,speed_ms,0,blend_radius_m)
  movel([0.309423, -1.280123, -2.629827, -0.802439, 1.570796, 1.880220],accel_mss,speed_ms,0,blend_radius_m)
  movel([0.307516, -1.286424, -2.626194, -0.799771, 1.570796, 1.878312],accel_mss,speed_ms,0,blend_radius_m)
  movel([0.305463, -1.292697, -2.622527, -0.797165, 1.570796, 1.876259],accel_mss,speed_ms,0,blend_radius_m)
  movel([0.297082, -1.317165, -2.607740, -0.787484, 1.570796, 1.867879],accel_mss,speed_ms,0,blend_radius_m)
  movel([0.293401, -1.328934, -2.600348, -0.783107, 1.570796, 1.864198],accel_mss,speed_ms,0,blend_radius_m)
  movel([0.291765, -1.334720, -2.596646, -0.781023, 1.570796, 1.862561],accel_mss,speed_ms,0,blend_radius_m)
  movel([0.290327, -1.340415, -2.592957, -0.779017, 1.570796, 1.861124],accel_mss,speed_ms,0,blend_radius_m)
  movel([0.289130, -1.346010, -2.589291, -0.777088, 1.570796, 1.859926],accel_mss,speed_ms,0,blend_radius_m)
  movel([0.288216, -1.351488, -2.585659, -0.775242, 1.570796, 1.859013],accel_mss,speed_ms,0,blend_radius_m)
  movel([0.287624, -1.356839, -2.582072, -0.773478, 1.570796, 1.858420],accel_mss,speed_ms,0,blend_radius_m)
  movel([0.287400, -1.362048, -2.578541, -0.771799, 1.570796, 1.858196],accel_mss,speed_ms,0,blend_radius_m)
  movel([0.287460, -1.364020, -2.577195, -0.771174, 1.570796, 1.858256],accel_mss,speed_ms,0,blend_radius_m)
  movel([0.287768, -1.365876, -2.575923, -0.770590, 1.570796, 1.858564],accel_mss,speed_ms,0,blend_radius_m)
  movel([0.288464, -1.367462, -2.574832, -0.770095, 1.570796, 1.859261],accel_mss,speed_ms,0,blend_radius_m)
  movel([0.289003, -1.368105, -2.574388, -0.769895, 1.570796, 1.859800],accel_mss,speed_ms,0,blend_radius_m)
  movel([0.289696, -1.368622, -2.574032, -0.769735, 1.570796, 1.860493],accel_mss,speed_ms,0,blend_radius_m)
  speed_ms = 0.005
  movel([0.289696, -1.359981, -2.569966, -0.782442, 1.570796, 1.860493],accel_mss,speed_ms,0,blend_radius_m)
  speed_ms = 0.040
  movel([0.277835, -1.333189, -2.587740, -0.791460, 1.570796, 1.848632],accel_mss,speed_ms,0,blend_radius_m)
  speed_ms = 0.005
  movel([0.277835, -1.342001, -2.591923, -0.778466, 1.570796, 1.848632],accel_mss,speed_ms,0,blend_radius_m)
  speed_ms = 0.025
  movel([0.277179, -1.342644, -2.591502, -0.778243, 1.570796, 1.847976],accel_mss,speed_ms,0,blend_radius_m)
  movel([0.276647, -1.343383, -2.591018, -0.777988, 1.570796, 1.847443],accel_mss,speed_ms,0,blend_radius_m)
  movel([0.276232, -1.344198, -2.590483, -0.777708, 1.570796, 1.847028],accel_mss,speed_ms,0,blend_radius_m)
  movel([0.275912, -1.345082, -2.589902, -0.777405, 1.570796, 1.846708],accel_mss,speed_ms,0,blend_radius_m)
  movel([0.275519, -1.346995, -2.588641, -0.776753, 1.570796, 1.846315],accel_mss,speed_ms,0,blend_radius_m)
  movel([0.275360, -1.349016, -2.587303, -0.776070, 1.570796, 1.846156],accel_mss,speed_ms,0,blend_radius_m)
  movel([0.275219, -1.354707, -2.583506, -0.774176, 1.570796, 1.846016],accel_mss,speed_ms,0,blend_radius_m)
  movel([0.274930, -1.356141, -2.582542, -0.773706, 1.570796, 1.845726],accel_mss,speed_ms,0,blend_radius_m)
  movel([0.274604, -1.356753, -2.582130, -0.773506, 1.570796, 1.845400],accel_mss,speed_ms,0,blend_radius_m)
  movel([0.274125, -1.357166, -2.581852, -0.773372, 1.570796, 1.844921],accel_mss,speed_ms,0,blend_radius_m)
  movel([0.273699, -1.357336, -2.581736, -0.773316, 1.570796, 1.844495],accel_mss,speed_ms,0,blend_radius_m)
  movel([0.273323, -1.357293, -2.581766, -0.773330, 1.570796, 1.844119],accel_mss,speed_ms,0,blend_radius_m)
  movel([0.272992, -1.357067, -2.581918, -0.773404, 1.570796, 1.843788],accel_mss,speed_ms,0,blend_radius_m)
  movel([0.272459, -1.356171, -2.582522, -0.773696, 1.570796, 1.843255],accel_mss,speed_ms,0,blend_radius_m)
  movel([0.272077, -1.354880, -2.583390, -0.774119, 1.570796, 1.842873],accel_mss,speed_ms,0,blend_radius_m)
  movel([0.271679, -1.352019, -2.585305, -0.775065, 1.570796, 1.842475],accel_mss,speed_ms,0,blend_radius_m)
  movel([0.271639, -1.350322, -2.586435, -0.775631, 1.570796, 1.842435],accel_mss,speed_ms,0,blend_radius_m)
  movel([0.270523, -1.352688, -2.584858, -0.774843, 1.570796, 1.841319],accel_mss,speed_ms,0,blend_radius_m)
  movel([0.269741, -1.355044, -2.583280, -0.774065, 1.570796, 1.840537],accel_mss,speed_ms,0,blend_radius_m)
  movel([0.269247, -1.357377, -2.581709, -0.773303, 1.570796, 1.840043],accel_mss,speed_ms,0,blend_radius_m)
  movel([0.269003, -1.359664, -2.580162, -0.772563, 1.570796, 1.839800],accel_mss,speed_ms,0,blend_radius_m)
  movel([0.268962, -1.361896, -2.578645, -0.771848, 1.570796, 1.839758],accel_mss,speed_ms,0,blend_radius_m)
  movel([0.269088, -1.364048, -2.577176, -0.771165, 1.570796, 1.839884],accel_mss,speed_ms,0,blend_radius_m)
  movel([0.269662, -1.368054, -2.574424, -0.769911, 1.570796, 1.840459],accel_mss,speed_ms,0,blend_radius_m)
  movel([0.269582, -1.368889, -2.573847, -0.769653, 1.570796, 1.840378],accel_mss,speed_ms,0,blend_radius_m)
  movel([0.269352, -1.369265, -2.573587, -0.769537, 1.570796, 1.840148],accel_mss,speed_ms,0,blend_radius_m)
  movel([0.268977, -1.369487, -2.573433, -0.769468, 1.570796, 1.839773],accel_mss,speed_ms,0,blend_radius_m)
  movel([0.268539, -1.369456, -2.573455, -0.769478, 1.570796, 1.839335],accel_mss,speed_ms,0,blend_radius_m)
  movel([0.267638, -1.369060, -2.573729, -0.769600, 1.570796, 1.838435],accel_mss,speed_ms,0,blend_radius_m)
  movel([0.266917, -1.368488, -2.574124, -0.769777, 1.570796, 1.837714],accel_mss,speed_ms,0,blend_radius_m)
  movel([0.266353, -1.367769, -2.574620, -0.770000, 1.570796, 1.837149],accel_mss,speed_ms,0,blend_radius_m)
  movel([0.265932, -1.366925, -2.575202, -0.770262, 1.570796, 1.836729],accel_mss,speed_ms,0,blend_radius_m)
  movel([0.265449, -1.364973, -2.576542, -0.770874, 1.570796, 1.836246],accel_mss,speed_ms,0,blend_radius_m)
  movel([0.265328, -1.362843, -2.577999, -0.771547, 1.570796, 1.836124],accel_mss,speed_ms,0,blend_radius_m)
  movel([0.264379, -1.367062, -2.575107, -0.770220, 1.570796, 1.835175],accel_mss,speed_ms,0,blend_radius_m)
  movel([0.264126, -1.369095, -2.573705, -0.769589, 1.570796, 1.834922],accel_mss,speed_ms,0,blend_radius_m)
  movel([0.264144, -1.371049, -2.572351, -0.768989, 1.570796, 1.834941],accel_mss,speed_ms,0,blend_radius_m)
  movel([0.264513, -1.372606, -2.571269, -0.768514, 1.570796, 1.835309],accel_mss,speed_ms,0,blend_radius_m)
  movel([0.265710, -1.375319, -2.569375, -0.767695, 1.570796, 1.836506],accel_mss,speed_ms,0,blend_radius_m)
  movel([0.266043, -1.376836, -2.568311, -0.767242, 1.570796, 1.836840],accel_mss,speed_ms,0,blend_radius_m)
  movel([0.266041, -1.377170, -2.568077, -0.767143, 1.570796, 1.836837],accel_mss,speed_ms,0,blend_radius_m)
  movel([0.265902, -1.377518, -2.567832, -0.767039, 1.570796, 1.836698],accel_mss,speed_ms,0,blend_radius_m)
  movel([0.265563, -1.377789, -2.567641, -0.766959, 1.570796, 1.836359],accel_mss,speed_ms,0,blend_radius_m)
  movel([0.265037, -1.377943, -2.567532, -0.766913, 1.570796, 1.835833],accel_mss,speed_ms,0,blend_radius_m)
  movel([0.263678, -1.378001, -2.567492, -0.766896, 1.570796, 1.834474],accel_mss,speed_ms,0,blend_radius_m)
  movel([0.261481, -1.377740, -2.567676, -0.766973, 1.570796, 1.832277],accel_mss,speed_ms,0,blend_radius_m)
  movel([0.261576, -1.378980, -2.566802, -0.766607, 1.570796, 1.832373],accel_mss,speed_ms,0,blend_radius_m)
  movel([0.261814, -1.380378, -2.565815, -0.766196, 1.570796, 1.832610],accel_mss,speed_ms,0,blend_radius_m)
  movel([0.262249, -1.381868, -2.564759, -0.765762, 1.570796, 1.833046],accel_mss,speed_ms,0,blend_radius_m)
  movel([0.262942, -1.383388, -2.563679, -0.765322, 1.570796, 1.833738],accel_mss,speed_ms,0,blend_radius_m)
  movel([0.265290, -1.385721, -2.562015, -0.764653, 1.570796, 1.836086],accel_mss,speed_ms,0,blend_radius_m)
  movel([0.266576, -1.387087, -2.561037, -0.764265, 1.570796, 1.837372],accel_mss,speed_ms,0,blend_radius_m)
  movel([0.266919, -1.387639, -2.560641, -0.764109, 1.570796, 1.837716],accel_mss,speed_ms,0,blend_radius_m)
  movel([0.266940, -1.388038, -2.560355, -0.763997, 1.570796, 1.837736],accel_mss,speed_ms,0,blend_radius_m)
  movel([0.266678, -1.388364, -2.560120, -0.763905, 1.570796, 1.837475],accel_mss,speed_ms,0,blend_radius_m)
  movel([0.266328, -1.388625, -2.559933, -0.763831, 1.570796, 1.837125],accel_mss,speed_ms,0,blend_radius_m)
  movel([0.265540, -1.388904, -2.559732, -0.763753, 1.570796, 1.836336],accel_mss,speed_ms,0,blend_radius_m)
  movel([0.264929, -1.388895, -2.559739, -0.763756, 1.570796, 1.835726],accel_mss,speed_ms,0,blend_radius_m)
  movel([0.264343, -1.388766, -2.559831, -0.763792, 1.570796, 1.835139],accel_mss,speed_ms,0,blend_radius_m)
  movel([0.263250, -1.388427, -2.560075, -0.763887, 1.570796, 1.834046],accel_mss,speed_ms,0,blend_radius_m)
  movel([0.263440, -1.390109, -2.558864, -0.763416, 1.570796, 1.834236],accel_mss,speed_ms,0,blend_radius_m)
  movel([0.263777, -1.391720, -2.557700, -0.762969, 1.570796, 1.834573],accel_mss,speed_ms,0,blend_radius_m)
  movel([0.264260, -1.393250, -2.556591, -0.762548, 1.570796, 1.835057],accel_mss,speed_ms,0,blend_radius_m)
  movel([0.264880, -1.394697, -2.555539, -0.762153, 1.570796, 1.835677],accel_mss,speed_ms,0,blend_radius_m)
  movel([0.265707, -1.395981, -2.554603, -0.761805, 1.570796, 1.836503],accel_mss,speed_ms,0,blend_radius_m)
  movel([0.266761, -1.397085, -2.553796, -0.761507, 1.570796, 1.837557],accel_mss,speed_ms,0,blend_radius_m)
  movel([0.269174, -1.399014, -2.552383, -0.760992, 1.570796, 1.839970],accel_mss,speed_ms,0,blend_radius_m)
  movel([0.269753, -1.399682, -2.551892, -0.760815, 1.570796, 1.840549],accel_mss,speed_ms,0,blend_radius_m)
  movel([0.269829, -1.400111, -2.551577, -0.760701, 1.570796, 1.840625],accel_mss,speed_ms,0,blend_radius_m)
  movel([0.269646, -1.400593, -2.551222, -0.760574, 1.570796, 1.840443],accel_mss,speed_ms,0,blend_radius_m)
  movel([0.269284, -1.400971, -2.550943, -0.760475, 1.570796, 1.840081],accel_mss,speed_ms,0,blend_radius_m)
  movel([0.268824, -1.401239, -2.550745, -0.760404, 1.570796, 1.839620],accel_mss,speed_ms,0,blend_radius_m)
  movel([0.267809, -1.401524, -2.550535, -0.760329, 1.570796, 1.838606],accel_mss,speed_ms,0,blend_radius_m)
  movel([0.266514, -1.401648, -2.550444, -0.760297, 1.570796, 1.837310],accel_mss,speed_ms,0,blend_radius_m)
  movel([0.265293, -1.401620, -2.550465, -0.760304, 1.570796, 1.836090],accel_mss,speed_ms,0,blend_radius_m)
  movel([0.264137, -1.401463, -2.550580, -0.760345, 1.570796, 1.834933],accel_mss,speed_ms,0,blend_radius_m)
  movel([0.263040, -1.401194, -2.550779, -0.760416, 1.570796, 1.833837],accel_mss,speed_ms,0,blend_radius_m)
  movel([0.263514, -1.402510, -2.549807, -0.760072, 1.570796, 1.834310],accel_mss,speed_ms,0,blend_radius_m)
  movel([0.264161, -1.403705, -2.548922, -0.759761, 1.570796, 1.834957],accel_mss,speed_ms,0,blend_radius_m)
  movel([0.264982, -1.404754, -2.548144, -0.759490, 1.570796, 1.835778],accel_mss,speed_ms,0,blend_radius_m)
  movel([0.265975, -1.405638, -2.547488, -0.759264, 1.570796, 1.836772],accel_mss,speed_ms,0,blend_radius_m)
  movel([0.267146, -1.406334, -2.546969, -0.759086, 1.570796, 1.837942],accel_mss,speed_ms,0,blend_radius_m)
  movel([0.268496, -1.406822, -2.546606, -0.758961, 1.570796, 1.839292],accel_mss,speed_ms,0,blend_radius_m)
  movel([0.270025, -1.407078, -2.546414, -0.758896, 1.570796, 1.840822],accel_mss,speed_ms,0,blend_radius_m)
  movel([0.271739, -1.407084, -2.546410, -0.758895, 1.570796, 1.842536],accel_mss,speed_ms,0,blend_radius_m)
  speed_ms = 0.005
  movel([0.271739, -1.398707, -2.542511, -0.771171, 1.570796, 1.842536],accel_mss,speed_ms,0,blend_radius_m)
  speed_ms = 0.040
  movel([0.280294, -1.390473, -2.548527, -0.773389, 1.570796, 1.851091],accel_mss,speed_ms,0,blend_radius_m)
  speed_ms = 0.005
  movel([0.280294, -1.398907, -2.552461, -0.761020, 1.570796, 1.851091],accel_mss,speed_ms,0,blend_radius_m)
  speed_ms = 0.025
  movel([0.277366, -1.397434, -2.553541, -0.761414, 1.570796, 1.848162],accel_mss,speed_ms,0,blend_radius_m)
  movel([0.276144, -1.396654, -2.554112, -0.761623, 1.570796, 1.846940],accel_mss,speed_ms,0,blend_radius_m)
  movel([0.275081, -1.395790, -2.554743, -0.761856, 1.570796, 1.845877],accel_mss,speed_ms,0,blend_radius_m)
  movel([0.274173, -1.394798, -2.555466, -0.762125, 1.570796, 1.844969],accel_mss,speed_ms,0,blend_radius_m)
  movel([0.273419, -1.393636, -2.556311, -0.762442, 1.570796, 1.844215],accel_mss,speed_ms,0,blend_radius_m)
  movel([0.272812, -1.392264, -2.557306, -0.762819, 1.570796, 1.843608],accel_mss,speed_ms,0,blend_radius_m)
  movel([0.272354, -1.390637, -2.558483, -0.763269, 1.570796, 1.843151],accel_mss,speed_ms,0,blend_radius_m)
  movel([0.271795, -1.387043, -2.561068, -0.764277, 1.570796, 1.842591],accel_mss,speed_ms,0,blend_radius_m)
  movel([0.271611, -1.383270, -2.563763, -0.765356, 1.570796, 1.842408],accel_mss,speed_ms,0,blend_radius_m)
  movel([0.271766, -1.379349, -2.566541, -0.766498, 1.570796, 1.842562],accel_mss,speed_ms,0,blend_radius_m)
  movel([0.272215, -1.375320, -2.569374, -0.767695, 1.570796, 1.843012],accel_mss,speed_ms,0,blend_radius_m)
  movel([0.272795, -1.371953, -2.571724, -0.768713, 1.570796, 1.843592],accel_mss,speed_ms,0,blend_radius_m)
  movel([0.273544, -1.368535, -2.574092, -0.769762, 1.570796, 1.844341],accel_mss,speed_ms,0,blend_radius_m)
  movel([0.275421, -1.361567, -2.578869, -0.771953, 1.570796, 1.846218],accel_mss,speed_ms,0,blend_radius_m)
  movel([0.282766, -1.337011, -2.595167, -0.780211, 1.570796, 1.853563],accel_mss,speed_ms,0,blend_radius_m)
  movel([0.284300, -1.331746, -2.598554, -0.782089, 1.570796, 1.855096],accel_mss,speed_ms,0,blend_radius_m)
  movel([0.285740, -1.326447, -2.601925, -0.784016, 1.570796, 1.856536],accel_mss,speed_ms,0,blend_radius_m)
  movel([0.287008, -1.321152, -2.605257, -0.785980, 1.570796, 1.857805],accel_mss,speed_ms,0,blend_radius_m)
  movel([0.288023, -1.315889, -2.608531, -0.787969, 1.570796, 1.858820],accel_mss,speed_ms,0,blend_radius_m)
  movel([0.288705, -1.310696, -2.611726, -0.789967, 1.570796, 1.859502],accel_mss,speed_ms,0,blend_radius_m)
  movel([0.288970, -1.305610, -2.614821, -0.791959, 1.570796, 1.859766],accel_mss,speed_ms,0,blend_radius_m)
  movel([0.288869, -1.301992, -2.617001, -0.793396, 1.570796, 1.859666],accel_mss,speed_ms,0,blend_radius_m)
  movel([0.288513, -1.298366, -2.619170, -0.794853, 1.570796, 1.859310],accel_mss,speed_ms,0,blend_radius_m)
  movel([0.287874, -1.294804, -2.621284, -0.796301, 1.570796, 1.858671],accel_mss,speed_ms,0,blend_radius_m)
  movel([0.286923, -1.291375, -2.623304, -0.797710, 1.570796, 1.857719],accel_mss,speed_ms,0,blend_radius_m)
  movel([0.285635, -1.288153, -2.625188, -0.799048, 1.570796, 1.856431],accel_mss,speed_ms,0,blend_radius_m)
  movel([0.283984, -1.285209, -2.626898, -0.800282, 1.570796, 1.854781],accel_mss,speed_ms,0,blend_radius_m)
  movel([0.281941, -1.282623, -2.628392, -0.801375, 1.570796, 1.852738],accel_mss,speed_ms,0,blend_radius_m)
  movel([0.279486, -1.280469, -2.629629, -0.802291, 1.570796, 1.850282],accel_mss,speed_ms,0,blend_radius_m)
  movel([0.278166, -1.279649, -2.630098, -0.802642, 1.570796, 1.848963],accel_mss,speed_ms,0,blend_radius_m)
  movel([0.276709, -1.278979, -2.630481, -0.802929, 1.570796, 1.847506],accel_mss,speed_ms,0,blend_radius_m)
  movel([0.275123, -1.278478, -2.630767, -0.803144, 1.570796, 1.845920],accel_mss,speed_ms,0,blend_radius_m)
  movel([0.273421, -1.278166, -2.630945, -0.803278, 1.570796, 1.844218],accel_mss,speed_ms,0,blend_radius_m)
  movel([0.271619, -1.278055, -2.631008, -0.803325, 1.570796, 1.842415],accel_mss,speed_ms,0,blend_radius_m)
  movel([0.269720, -1.278167, -2.630945, -0.803277, 1.570796, 1.840517],accel_mss,speed_ms,0,blend_radius_m)
  movel([0.267745, -1.278513, -2.630747, -0.803129, 1.570796, 1.838541],accel_mss,speed_ms,0,blend_radius_m)
  movel([0.265704, -1.279113, -2.630405, -0.802871, 1.570796, 1.836500],accel_mss,speed_ms,0,blend_radius_m)
  speed_ms = 0.005
  movel([0.265704, -1.269944, -2.625941, -0.816505, 1.570796, 1.836500],accel_mss,speed_ms,0,blend_radius_m)
  speed_ms = 0.040
  movel([0.261221, -1.258722, -2.632193, -0.821474, 1.570796, 1.832018],accel_mss,speed_ms,0,blend_radius_m)
  speed_ms = 0.005
  movel([0.261221, -1.267947, -2.636707, -0.807735, 1.570796, 1.832018],accel_mss,speed_ms,0,blend_radius_m)
  speed_ms = 0.025
  movel([0.261256, -1.266555, -2.637482, -0.808352, 1.570796, 1.832052],accel_mss,speed_ms,0,blend_radius_m)
  movel([0.261456, -1.265113, -2.638282, -0.808994, 1.570796, 1.832252],accel_mss,speed_ms,0,blend_radius_m)
  movel([0.262252, -1.262120, -2.639935, -0.810334, 1.570796, 1.833048],accel_mss,speed_ms,0,blend_radius_m)
  movel([0.263426, -1.259032, -2.641629, -0.811728, 1.570796, 1.834222],accel_mss,speed_ms,0,blend_radius_m)
  movel([0.264782, -1.255927, -2.643320, -0.813141, 1.570796, 1.835578],accel_mss,speed_ms,0,blend_radius_m)
  speed_ms = 0.005
  movel([0.264782, -1.246646, -2.638752, -0.826991, 1.570796, 1.835578],accel_mss,speed_ms,0,blend_radius_m)
  speed_ms = 0.040
  movel([0.268657, -1.247900, -2.638079, -0.826410, 1.570796, 1.839454],accel_mss,speed_ms,0,blend_radius_m)
  speed_ms = 0.005
  movel([0.268657, -1.257176, -2.642642, -0.812572, 1.570796, 1.839454],accel_mss,speed_ms,0,blend_radius_m)
  speed_ms = 0.025
  movel([0.268335, -1.256049, -2.643254, -0.813086, 1.570796, 1.839131],accel_mss,speed_ms,0,blend_radius_m)
  movel([0.268177, -1.254867, -2.643895, -0.813627, 1.570796, 1.838973],accel_mss,speed_ms,0,blend_radius_m)
  movel([0.268308, -1.252352, -2.645254, -0.814783, 1.570796, 1.839104],accel_mss,speed_ms,0,blend_radius_m)
  movel([0.268970, -1.249683, -2.646687, -0.816019, 1.570796, 1.839766],accel_mss,speed_ms,0,blend_radius_m)
  movel([0.270079, -1.246903, -2.648171, -0.817315, 1.570796, 1.840875],accel_mss,speed_ms,0,blend_radius_m)
  movel([0.271549, -1.244063, -2.649677, -0.818649, 1.570796, 1.842345],accel_mss,speed_ms,0,blend_radius_m)
  movel([0.273295, -1.241214, -2.651179, -0.819997, 1.570796, 1.844091],accel_mss,speed_ms,0,blend_radius_m)
  movel([0.275228, -1.238405, -2.652650, -0.821334, 1.570796, 1.846024],accel_mss,speed_ms,0,blend_radius_m)
  movel([0.277259, -1.235691, -2.654062, -0.822635, 1.570796, 1.848055],accel_mss,speed_ms,0,blend_radius_m)
  speed_ms = 0.005
  movel([0.277259, -1.226322, -2.649402, -0.836665, 1.570796, 1.848055],accel_mss,speed_ms,0,blend_radius_m)
  speed_ms = 0.040
  movel([0.300694, -1.205116, -2.660011, -0.847262, 1.570796, 1.871491],accel_mss,speed_ms,0,blend_radius_m)
  speed_ms = 0.005
  movel([0.300694, -1.214566, -2.664767, -0.833056, 1.570796, 1.871491],accel_mss,speed_ms,0,blend_radius_m)
  speed_ms = 0.025
  movel([0.298485, -1.215961, -2.664075, -0.832352, 1.570796, 1.869281],accel_mss,speed_ms,0,blend_radius_m)
  movel([0.296248, -1.217535, -2.663293, -0.831561, 1.570796, 1.867044],accel_mss,speed_ms,0,blend_radius_m)
  movel([0.294018, -1.219262, -2.662432, -0.830696, 1.570796, 1.864814],accel_mss,speed_ms,0,blend_radius_m)
  movel([0.291822, -1.221122, -2.661499, -0.829768, 1.570796, 1.862618],accel_mss,speed_ms,0,blend_radius_m)
  movel([0.289695, -1.223097, -2.660506, -0.828787, 1.570796, 1.860491],accel_mss,speed_ms,0,blend_radius_m)
  movel([0.287667, -1.225159, -2.659463, -0.827767, 1.570796, 1.858464],accel_mss,speed_ms,0,blend_radius_m)
  movel([0.285770, -1.227294, -2.658379, -0.826716, 1.570796, 1.856566],accel_mss,speed_ms,0,blend_radius_m)
  movel([0.284034, -1.229480, -2.657263, -0.825646, 1.570796, 1.854830],accel_mss,speed_ms,0,blend_radius_m)
  movel([0.282489, -1.231693, -2.656128, -0.824569, 1.570796, 1.853285],accel_mss,speed_ms,0,blend_radius_m)
  movel([0.281163, -1.233916, -2.654981, -0.823491, 1.570796, 1.851959],accel_mss,speed_ms,0,blend_radius_m)
  movel([0.280085, -1.236129, -2.653835, -0.822425, 1.570796, 1.850882],accel_mss,speed_ms,0,blend_radius_m)
  movel([0.279284, -1.238313, -2.652698, -0.821378, 1.570796, 1.850081],accel_mss,speed_ms,0,blend_radius_m)
  movel([0.278791, -1.240447, -2.651581, -0.820361, 1.570796, 1.849587],accel_mss,speed_ms,0,blend_radius_m)
  movel([0.278632, -1.242515, -2.650494, -0.819380, 1.570796, 1.849428],accel_mss,speed_ms,0,blend_radius_m)
  movel([0.278831, -1.244499, -2.649447, -0.818444, 1.570796, 1.849627],accel_mss,speed_ms,0,blend_radius_m)
  movel([0.279419, -1.246382, -2.648448, -0.817559, 1.570796, 1.850216],accel_mss,speed_ms,0,blend_radius_m)
  speed_ms = 0.005
  movel([0.279419, -1.237058, -2.643836, -0.831495, 1.570796, 1.850216],accel_mss,speed_ms,0,blend_radius_m)
  speed_ms = 0.040
  movel([0.289856, -1.230979, -2.647004, -0.834406, 1.570796, 1.860653],accel_mss,speed_ms,0,blend_radius_m)
  speed_ms = 0.005
  movel([0.289856, -1.240329, -2.651643, -0.820417, 1.570796, 1.860653],accel_mss,speed_ms,0,blend_radius_m)
  speed_ms = 0.025
  movel([0.289896, -1.238660, -2.652517, -0.821212, 1.570796, 1.860692],accel_mss,speed_ms,0,blend_radius_m)
  movel([0.290100, -1.236921, -2.653423, -0.822045, 1.570796, 1.860896],accel_mss,speed_ms,0,blend_radius_m)
  movel([0.290464, -1.235132, -2.654352, -0.822905, 1.570796, 1.861260],accel_mss,speed_ms,0,blend_radius_m)
  movel([0.290984, -1.233303, -2.655298, -0.823788, 1.570796, 1.861781],accel_mss,speed_ms,0,blend_radius_m)
  movel([0.291655, -1.231451, -2.656252, -0.824686, 1.570796, 1.862451],accel_mss,speed_ms,0,blend_radius_m)
  movel([0.292475, -1.229590, -2.657206, -0.825592, 1.570796, 1.863271],accel_mss,speed_ms,0,blend_radius_m)
  movel([0.293441, -1.227732, -2.658156, -0.826502, 1.570796, 1.864238],accel_mss,speed_ms,0,blend_radius_m)
  movel([0.294546, -1.225896, -2.659090, -0.827404, 1.570796, 1.865343],accel_mss,speed_ms,0,blend_radius_m)
  movel([0.295787, -1.224094, -2.660002, -0.828293, 1.570796, 1.866583],accel_mss,speed_ms,0,blend_radius_m)
  movel([0.297162, -1.222342, -2.660886, -0.829161, 1.570796, 1.867958],accel_mss,speed_ms,0,blend_radius_m)
  movel([0.298659, -1.220662, -2.661730, -0.829997, 1.570796, 1.869455],accel_mss,speed_ms,0,blend_radius_m)
  movel([0.300282, -1.219061, -2.662532, -0.830796, 1.570796, 1.871079],accel_mss,speed_ms,0,blend_radius_m)
  movel([0.302023, -1.217559, -2.663281, -0.831549, 1.570796, 1.872819],accel_mss,speed_ms,0,blend_radius_m)
  movel([0.303876, -1.216172, -2.663971, -0.832246, 1.570796, 1.874673],accel_mss,speed_ms,0,blend_radius_m)
  movel([0.305836, -1.214918, -2.664592, -0.832878, 1.570796, 1.876632],accel_mss,speed_ms,0,blend_radius_m)
  movel([0.307895, -1.213813, -2.665139, -0.833437, 1.570796, 1.878691],accel_mss,speed_ms,0,blend_radius_m)
  movel([0.309920, -1.212937, -2.665571, -0.833881, 1.570796, 1.880716],accel_mss,speed_ms,0,blend_radius_m)
  movel([0.311897, -1.212287, -2.665891, -0.834211, 1.570796, 1.882693],accel_mss,speed_ms,0,blend_radius_m)
  movel([0.313815, -1.211854, -2.666104, -0.834431, 1.570796, 1.884612],accel_mss,speed_ms,0,blend_radius_m)
  movel([0.315670, -1.211629, -2.666215, -0.834545, 1.570796, 1.886466],accel_mss,speed_ms,0,blend_radius_m)
  movel([0.317450, -1.211601, -2.666228, -0.834559, 1.570796, 1.888247],accel_mss,speed_ms,0,blend_radius_m)
  movel([0.319144, -1.211765, -2.666148, -0.834476, 1.570796, 1.889940],accel_mss,speed_ms,0,blend_radius_m)
  movel([0.320749, -1.212102, -2.665982, -0.834305, 1.570796, 1.891546],accel_mss,speed_ms,0,blend_radius_m)
  movel([0.322249, -1.212608, -2.665733, -0.834048, 1.570796, 1.893046],accel_mss,speed_ms,0,blend_radius_m)
  movel([0.323641, -1.213270, -2.665407, -0.833712, 1.570796, 1.894437],accel_mss,speed_ms,0,blend_radius_m)
  movel([0.326068, -1.215016, -2.664544, -0.832829, 1.570796, 1.896865],accel_mss,speed_ms,0,blend_radius_m)
  movel([0.327083, -1.216078, -2.664017, -0.832293, 1.570796, 1.897880],accel_mss,speed_ms,0,blend_radius_m)
  movel([0.328692, -1.218523, -2.662801, -0.831066, 1.570796, 1.899488],accel_mss,speed_ms,0,blend_radius_m)
  movel([0.329269, -1.219881, -2.662122, -0.830387, 1.570796, 1.900065],accel_mss,speed_ms,0,blend_radius_m)
  movel([0.329683, -1.221315, -2.661402, -0.829671, 1.570796, 1.900479],accel_mss,speed_ms,0,blend_radius_m)
  speed_ms = 0.005
  movel([0.329683, -1.211889, -2.656677, -0.843822, 1.570796, 1.900479],accel_mss,speed_ms,0,blend_radius_m)
  speed_ms = 0.040
  movel([0.334756, -1.223526, -2.650830, -0.838033, 1.570796, 1.905552],accel_mss,speed_ms,0,blend_radius_m)
  speed_ms = 0.005
  movel([0.334756, -1.232907, -2.655503, -0.823980, 1.570796, 1.905552],accel_mss,speed_ms,0,blend_radius_m)
  speed_ms = 0.025
  movel([0.334182, -1.230721, -2.656627, -0.825041, 1.570796, 1.904978],accel_mss,speed_ms,0,blend_radius_m)
  movel([0.333230, -1.228813, -2.657604, -0.825972, 1.570796, 1.904027],accel_mss,speed_ms,0,blend_radius_m)
  movel([0.331927, -1.227205, -2.658424, -0.826760, 1.570796, 1.902723],accel_mss,speed_ms,0,blend_radius_m)
  movel([0.330293, -1.225916, -2.659079, -0.827394, 1.570796, 1.901089],accel_mss,speed_ms,0,blend_radius_m)
  movel([0.328362, -1.224966, -2.659561, -0.827862, 1.570796, 1.899158],accel_mss,speed_ms,0,blend_radius_m)
  movel([0.326156, -1.224377, -2.659859, -0.828153, 1.570796, 1.896952],accel_mss,speed_ms,0,blend_radius_m)
  movel([0.323707, -1.224166, -2.659966, -0.828257, 1.570796, 1.894504],accel_mss,speed_ms,0,blend_radius_m)
  movel([0.321041, -1.224350, -2.659873, -0.828166, 1.570796, 1.891837],accel_mss,speed_ms,0,blend_radius_m)
  movel([0.318195, -1.224946, -2.659571, -0.827872, 1.570796, 1.888991],accel_mss,speed_ms,0,blend_radius_m)
  movel([0.315229, -1.225952, -2.659061, -0.827376, 1.570796, 1.886025],accel_mss,speed_ms,0,blend_radius_m)
  movel([0.312254, -1.227344, -2.658353, -0.826692, 1.570796, 1.883050],accel_mss,speed_ms,0,blend_radius_m)
  movel([0.309387, -1.229098, -2.657458, -0.825833, 1.570796, 1.880183],accel_mss,speed_ms,0,blend_radius_m)
  movel([0.306734, -1.231194, -2.656384, -0.824811, 1.570796, 1.877531],accel_mss,speed_ms,0,blend_radius_m)
  movel([0.305526, -1.232362, -2.655783, -0.824244, 1.570796, 1.876323],accel_mss,speed_ms,0,blend_radius_m)
  movel([0.304412, -1.233603, -2.655144, -0.823643, 1.570796, 1.875209],accel_mss,speed_ms,0,blend_radius_m)
  movel([0.303406, -1.234916, -2.654464, -0.823009, 1.570796, 1.874202],accel_mss,speed_ms,0,blend_radius_m)
  movel([0.302523, -1.236303, -2.653745, -0.822342, 1.570796, 1.873320],accel_mss,speed_ms,0,blend_radius_m)
  movel([0.301774, -1.237753, -2.652990, -0.821646, 1.570796, 1.872570],accel_mss,speed_ms,0,blend_radius_m)
  movel([0.301178, -1.239264, -2.652201, -0.820924, 1.570796, 1.871974],accel_mss,speed_ms,0,blend_radius_m)
  speed_ms = 0.005
  movel([0.301178, -1.229910, -2.647557, -0.834922, 1.570796, 1.871974],accel_mss,speed_ms,0,blend_radius_m)
  speed_ms = 0.040
  movel([0.314688, -1.235201, -2.644808, -0.832380, 1.570796, 1.885485],accel_mss,speed_ms,0,blend_radius_m)
  speed_ms = 0.005
  movel([0.314688, -1.244533, -2.649428, -0.818427, 1.570796, 1.885485],accel_mss,speed_ms,0,blend_radius_m)
  speed_ms = 0.025
  movel([0.316787, -1.243271, -2.650096, -0.819023, 1.570796, 1.887583],accel_mss,speed_ms,0,blend_radius_m)
  movel([0.318910, -1.242297, -2.650609, -0.819483, 1.570796, 1.889706],accel_mss,speed_ms,0,blend_radius_m)
  movel([0.321030, -1.241601, -2.650975, -0.819813, 1.570796, 1.891826],accel_mss,speed_ms,0,blend_radius_m)
  movel([0.323108, -1.241174, -2.651200, -0.820015, 1.570796, 1.893904],accel_mss,speed_ms,0,blend_radius_m)
  movel([0.325112, -1.241002, -2.651290, -0.820097, 1.570796, 1.895908],accel_mss,speed_ms,0,blend_radius_m)
  movel([0.327006, -1.241070, -2.651255, -0.820065, 1.570796, 1.897802],accel_mss,speed_ms,0,blend_radius_m)
  movel([0.328762, -1.241365, -2.651099, -0.819925, 1.570796, 1.899558],accel_mss,speed_ms,0,blend_radius_m)
  movel([0.330341, -1.241872, -2.650833, -0.819684, 1.570796, 1.901137],accel_mss,speed_ms,0,blend_radius_m)
  movel([0.331962, -1.242808, -2.650340, -0.819241, 1.570796, 1.902758],accel_mss,speed_ms,0,blend_radius_m)
  movel([0.333078, -1.244035, -2.649692, -0.818662, 1.570796, 1.903875],accel_mss,speed_ms,0,blend_radius_m)
  movel([0.333747, -1.245520, -2.648905, -0.817963, 1.570796, 1.904543],accel_mss,speed_ms,0,blend_radius_m)
  movel([0.334013, -1.247232, -2.647995, -0.817161, 1.570796, 1.904809],accel_mss,speed_ms,0,blend_radius_m)
  movel([0.333931, -1.249132, -2.646982, -0.816275, 1.570796, 1.904727],accel_mss,speed_ms,0,blend_radius_m)
  movel([0.333551, -1.251192, -2.645878, -0.815320, 1.570796, 1.904347],accel_mss,speed_ms,0,blend_radius_m)
  movel([0.332923, -1.253376, -2.644701, -0.814311, 1.570796, 1.903720],accel_mss,speed_ms,0,blend_radius_m)
  movel([0.332103, -1.255654, -2.643469, -0.813266, 1.570796, 1.902899],accel_mss,speed_ms,0,blend_radius_m)
  speed_ms = 0.005
  movel([0.332103, -1.246371, -2.638899, -0.827119, 1.570796, 1.902899],accel_mss,speed_ms,0,blend_radius_m)
  speed_ms = 0.040
  movel([0.318559, -1.246626, -2.638762, -0.827001, 1.570796, 1.889356],accel_mss,speed_ms,0,blend_radius_m)
  speed_ms = 0.005
  movel([0.318559, -1.255908, -2.643331, -0.813150, 1.570796, 1.889356],accel_mss,speed_ms,0,blend_radius_m)
  speed_ms = 0.025
  movel([0.320362, -1.256055, -2.643251, -0.813083, 1.570796, 1.891158],accel_mss,speed_ms,0,blend_radius_m)
  movel([0.321966, -1.256425, -2.643050, -0.812914, 1.570796, 1.892763],accel_mss,speed_ms,0,blend_radius_m)
  movel([0.323375, -1.257010, -2.642732, -0.812647, 1.570796, 1.894171],accel_mss,speed_ms,0,blend_radius_m)
  movel([0.324594, -1.257786, -2.642309, -0.812294, 1.570796, 1.895390],accel_mss,speed_ms,0,blend_radius_m)
  movel([0.325628, -1.258740, -2.641789, -0.811861, 1.570796, 1.896424],accel_mss,speed_ms,0,blend_radius_m)
  movel([0.326481, -1.259853, -2.641180, -0.811356, 1.570796, 1.897278],accel_mss,speed_ms,0,blend_radius_m)
  movel([0.327161, -1.261109, -2.640491, -0.810789, 1.570796, 1.897957],accel_mss,speed_ms,0,blend_radius_m)
  movel([0.327667, -1.262494, -2.639729, -0.810166, 1.570796, 1.898464],accel_mss,speed_ms,0,blend_radius_m)
  movel([0.328012, -1.263990, -2.638903, -0.809495, 1.570796, 1.898808],accel_mss,speed_ms,0,blend_radius_m)
  movel([0.328198, -1.265580, -2.638023, -0.808785, 1.570796, 1.898994],accel_mss,speed_ms,0,blend_radius_m)
  movel([0.328228, -1.267249, -2.637096, -0.808044, 1.570796, 1.899025],accel_mss,speed_ms,0,blend_radius_m)
  movel([0.328113, -1.268980, -2.636130, -0.807278, 1.570796, 1.898909],accel_mss,speed_ms,0,blend_radius_m)
  movel([0.327854, -1.270759, -2.635134, -0.806495, 1.570796, 1.898650],accel_mss,speed_ms,0,blend_radius_m)
  movel([0.326930, -1.274395, -2.633087, -0.804908, 1.570796, 1.897726],accel_mss,speed_ms,0,blend_radius_m)
  movel([0.326274, -1.276224, -2.632050, -0.804115, 1.570796, 1.897070],accel_mss,speed_ms,0,blend_radius_m)
  movel([0.326267, -1.275642, -2.632380, -0.804367, 1.570796, 1.897063],accel_mss,speed_ms,0,blend_radius_m)
  speed_ms = 0.005
  movel([0.326267, -1.266455, -2.627901, -0.818033, 1.570796, 1.897063],accel_mss,speed_ms,0,blend_radius_m)
  speed_ms = 0.040
  movel([0.336306, -1.272774, -2.624340, -0.815276, 1.570796, 1.907103],accel_mss,speed_ms,0,blend_radius_m)
  speed_ms = 0.005
  movel([0.336306, -1.281929, -2.628791, -0.801669, 1.570796, 1.907103],accel_mss,speed_ms,0,blend_radius_m)
  speed_ms = 0.025
  movel([0.334244, -1.284171, -2.627498, -0.800719, 1.570796, 1.905040],accel_mss,speed_ms,0,blend_radius_m)
  movel([0.332389, -1.286519, -2.626139, -0.799731, 1.570796, 1.903186],accel_mss,speed_ms,0,blend_radius_m)
  movel([0.330700, -1.288929, -2.624736, -0.798724, 1.570796, 1.901497],accel_mss,speed_ms,0,blend_radius_m)
  movel([0.329130, -1.291361, -2.623312, -0.797716, 1.570796, 1.899926],accel_mss,speed_ms,0,blend_radius_m)
  movel([0.327524, -1.294055, -2.621727, -0.796608, 1.570796, 1.898320],accel_mss,speed_ms,0,blend_radius_m)
  movel([0.326844, -1.295404, -2.620929, -0.796056, 1.570796, 1.897640],accel_mss,speed_ms,0,blend_radius_m)
  movel([0.326299, -1.296748, -2.620132, -0.795509, 1.570796, 1.897096],accel_mss,speed_ms,0,blend_radius_m)
  movel([0.325926, -1.298077, -2.619342, -0.794970, 1.570796, 1.896722],accel_mss,speed_ms,0,blend_radius_m)
  movel([0.325769, -1.299349, -2.618584, -0.794456, 1.570796, 1.896566],accel_mss,speed_ms,0,blend_radius_m)
  movel([0.325872, -1.300505, -2.617893, -0.793991, 1.570796, 1.896669],accel_mss,speed_ms,0,blend_radius_m)
  movel([0.326269, -1.301494, -2.617300, -0.793595, 1.570796, 1.897065],accel_mss,speed_ms,0,blend_radius_m)
  movel([0.327365, -1.302700, -2.616576, -0.793113, 1.570796, 1.898161],accel_mss,speed_ms,0,blend_radius_m)
  movel([0.327903, -1.303303, -2.616213, -0.792873, 1.570796, 1.898700],accel_mss,speed_ms,0,blend_radius_m)
  movel([0.328285, -1.304021, -2.615781, -0.792588, 1.570796, 1.899081],accel_mss,speed_ms,0,blend_radius_m)
  movel([0.328394, -1.305055, -2.615156, -0.792178, 1.570796, 1.899190],accel_mss,speed_ms,0,blend_radius_m)
  movel([0.328181, -1.306307, -2.614398, -0.791684, 1.570796, 1.898977],accel_mss,speed_ms,0,blend_radius_m)
  movel([0.327719, -1.307711, -2.613546, -0.791132, 1.570796, 1.898515],accel_mss,speed_ms,0,blend_radius_m)
  movel([0.327078, -1.309199, -2.612640, -0.790550, 1.570796, 1.897874],accel_mss,speed_ms,0,blend_radius_m)
  movel([0.325533, -1.312163, -2.610827, -0.789399, 1.570796, 1.896329],accel_mss,speed_ms,0,blend_radius_m)
  movel([0.320752, -1.320285, -2.605798, -0.786305, 1.570796, 1.891548],accel_mss,speed_ms,0,blend_radius_m)
  movel([0.317462, -1.325853, -2.602301, -0.784235, 1.570796, 1.888258],accel_mss,speed_ms,0,blend_radius_m)
  movel([0.316573, -1.327574, -2.601212, -0.783603, 1.570796, 1.887369],accel_mss,speed_ms,0,blend_radius_m)
  movel([0.315744, -1.329422, -2.600038, -0.782930, 1.570796, 1.886541],accel_mss,speed_ms,0,blend_radius_m)
  movel([0.314354, -1.333338, -2.597534, -0.781517, 1.570796, 1.885150],accel_mss,speed_ms,0,blend_radius_m)
  movel([0.313837, -1.335328, -2.596254, -0.780807, 1.570796, 1.884633],accel_mss,speed_ms,0,blend_radius_m)
  movel([0.313467, -1.337286, -2.594989, -0.780114, 1.570796, 1.884264],accel_mss,speed_ms,0,blend_radius_m)
  movel([0.313266, -1.339173, -2.593766, -0.779450, 1.570796, 1.884062],accel_mss,speed_ms,0,blend_radius_m)
  movel([0.313253, -1.340953, -2.592607, -0.778829, 1.570796, 1.884050],accel_mss,speed_ms,0,blend_radius_m)
  movel([0.313452, -1.342583, -2.591542, -0.778264, 1.570796, 1.884249],accel_mss,speed_ms,0,blend_radius_m)
  movel([0.313880, -1.344033, -2.590592, -0.777765, 1.570796, 1.884677],accel_mss,speed_ms,0,blend_radius_m)
  movel([0.314563, -1.345260, -2.589785, -0.777344, 1.570796, 1.885359],accel_mss,speed_ms,0,blend_radius_m)
  movel([0.315519, -1.346229, -2.589146, -0.777014, 1.570796, 1.886315],accel_mss,speed_ms,0,blend_radius_m)
  movel([0.316768, -1.346905, -2.588701, -0.776784, 1.570796, 1.887564],accel_mss,speed_ms,0,blend_radius_m)
  movel([0.318335, -1.347248, -2.588474, -0.776667, 1.570796, 1.889132],accel_mss,speed_ms,0,blend_radius_m)
  movel([0.320242, -1.347225, -2.588489, -0.776675, 1.570796, 1.891038],accel_mss,speed_ms,0,blend_radius_m)
  movel([0.322513, -1.346797, -2.588772, -0.776821, 1.570796, 1.893309],accel_mss,speed_ms,0,blend_radius_m)
  movel([0.324337, -1.346218, -2.589154, -0.777017, 1.570796, 1.895133],accel_mss,speed_ms,0,blend_radius_m)
  movel([0.326152, -1.345465, -2.589650, -0.777274, 1.570796, 1.896948],accel_mss,speed_ms,0,blend_radius_m)
  movel([0.327962, -1.344564, -2.590242, -0.777582, 1.570796, 1.898758],accel_mss,speed_ms,0,blend_radius_m)
  movel([0.329764, -1.343545, -2.590912, -0.777933, 1.570796, 1.900560],accel_mss,speed_ms,0,blend_radius_m)
  movel([0.333342, -1.341268, -2.592401, -0.778720, 1.570796, 1.904138],accel_mss,speed_ms,0,blend_radius_m)
  movel([0.336882, -1.338869, -2.593963, -0.779557, 1.570796, 1.907679],accel_mss,speed_ms,0,blend_radius_m)
  movel([0.340490, -1.336543, -2.595470, -0.780376, 1.570796, 1.911286],accel_mss,speed_ms,0,blend_radius_m)
  movel([0.342340, -1.335471, -2.596162, -0.780756, 1.570796, 1.913136],accel_mss,speed_ms,0,blend_radius_m)
  movel([0.344201, -1.334508, -2.596782, -0.781099, 1.570796, 1.914997],accel_mss,speed_ms,0,blend_radius_m)
  movel([0.346059, -1.333687, -2.597310, -0.781392, 1.570796, 1.916855],accel_mss,speed_ms,0,blend_radius_m)
  movel([0.347899, -1.333045, -2.597722, -0.781622, 1.570796, 1.918695],accel_mss,speed_ms,0,blend_radius_m)
  movel([0.349702, -1.332616, -2.597997, -0.781776, 1.570796, 1.920498],accel_mss,speed_ms,0,blend_radius_m)
  movel([0.351457, -1.332438, -2.598111, -0.781840, 1.570796, 1.922253],accel_mss,speed_ms,0,blend_radius_m)
  movel([0.355050, -1.332648, -2.597977, -0.781764, 1.570796, 1.925847],accel_mss,speed_ms,0,blend_radius_m)
  movel([0.356286, -1.332624, -2.597992, -0.781773, 1.570796, 1.927083],accel_mss,speed_ms,0,blend_radius_m)
  movel([0.357621, -1.332385, -2.598145, -0.781859, 1.570796, 1.928417],accel_mss,speed_ms,0,blend_radius_m)
  movel([0.358994, -1.331881, -2.598468, -0.782040, 1.570796, 1.929790],accel_mss,speed_ms,0,blend_radius_m)
  movel([0.360280, -1.331108, -2.598962, -0.782319, 1.570796, 1.931076],accel_mss,speed_ms,0,blend_radius_m)
  movel([0.360854, -1.330617, -2.599276, -0.782496, 1.570796, 1.931650],accel_mss,speed_ms,0,blend_radius_m)
  movel([0.361360, -1.330056, -2.599634, -0.782699, 1.570796, 1.932157],accel_mss,speed_ms,0,blend_radius_m)
  speed_ms = 0.005
  movel([0.361360, -1.321171, -2.595398, -0.795820, 1.570796, 1.932157],accel_mss,speed_ms,0,blend_radius_m)
  speed_ms = 0.040
  movel([0.369046, -1.309954, -2.602373, -0.800062, 1.570796, 1.939842],accel_mss,speed_ms,0,blend_radius_m)
  speed_ms = 0.005
  movel([0.369046, -1.318906, -2.606659, -0.786825, 1.570796, 1.939842],accel_mss,speed_ms,0,blend_radius_m)
  speed_ms = 0.025
  movel([0.369408, -1.319136, -2.606515, -0.786738, 1.570796, 1.940204],accel_mss,speed_ms,0,blend_radius_m)
  movel([0.369364, -1.319664, -2.606186, -0.786539, 1.570796, 1.940160],accel_mss,speed_ms,0,blend_radius_m)
  movel([0.369004, -1.320281, -2.605801, -0.786307, 1.570796, 1.939801],accel_mss,speed_ms,0,blend_radius_m)
  movel([0.368431, -1.320783, -2.605487, -0.786118, 1.570796, 1.939228],accel_mss,speed_ms,0,blend_radius_m)
  movel([0.367782, -1.321068, -2.605310, -0.786012, 1.570796, 1.938579],accel_mss,speed_ms,0,blend_radius_m)
  movel([0.367136, -1.321214, -2.605218, -0.785957, 1.570796, 1.937932],accel_mss,speed_ms,0,blend_radius_m)
  movel([0.365854, -1.321367, -2.605122, -0.785900, 1.570796, 1.936650],accel_mss,speed_ms,0,blend_radius_m)
  movel([0.364910, -1.321584, -2.604986, -0.785819, 1.570796, 1.935707],accel_mss,speed_ms,0,blend_radius_m)
  movel([0.363963, -1.321933, -2.604768, -0.785688, 1.570796, 1.934759],accel_mss,speed_ms,0,blend_radius_m)
  movel([0.362069, -1.322937, -2.604138, -0.785314, 1.570796, 1.932865],accel_mss,speed_ms,0,blend_radius_m)
  movel([0.360207, -1.324222, -2.603330, -0.784837, 1.570796, 1.931004],accel_mss,speed_ms,0,blend_radius_m)
  movel([0.358417, -1.325615, -2.602452, -0.784323, 1.570796, 1.929214],accel_mss,speed_ms,0,blend_radius_m)
  movel([0.358005, -1.325979, -2.602221, -0.784188, 1.570796, 1.928801],accel_mss,speed_ms,0,blend_radius_m)
  movel([0.357731, -1.326388, -2.601963, -0.784038, 1.570796, 1.928528],accel_mss,speed_ms,0,blend_radius_m)
  movel([0.357770, -1.326812, -2.601695, -0.783883, 1.570796, 1.928566],accel_mss,speed_ms,0,blend_radius_m)
  movel([0.358082, -1.327090, -2.601519, -0.783781, 1.570796, 1.928878],accel_mss,speed_ms,0,blend_radius_m)
  movel([0.358950, -1.327508, -2.601254, -0.783627, 1.570796, 1.929747],accel_mss,speed_ms,0,blend_radius_m)
  movel([0.359935, -1.327765, -2.601090, -0.783533, 1.570796, 1.930731],accel_mss,speed_ms,0,blend_radius_m)
  movel([0.361017, -1.327868, -2.601025, -0.783496, 1.570796, 1.931813],accel_mss,speed_ms,0,blend_radius_m)
  movel([0.362176, -1.327814, -2.601060, -0.783516, 1.570796, 1.932972],accel_mss,speed_ms,0,blend_radius_m)
  movel([0.363384, -1.327611, -2.601188, -0.783590, 1.570796, 1.934181],accel_mss,speed_ms,0,blend_radius_m)
  movel([0.364625, -1.327256, -2.601413, -0.783720, 1.570796, 1.935421],accel_mss,speed_ms,0,blend_radius_m)
  movel([0.365872, -1.326755, -2.601730, -0.783903, 1.570796, 1.936669],accel_mss,speed_ms,0,blend_radius_m)
  movel([0.367107, -1.326107, -2.602141, -0.784141, 1.570796, 1.937904],accel_mss,speed_ms,0,blend_radius_m)
  movel([0.366838, -1.326772, -2.601720, -0.783897, 1.570796, 1.937634],accel_mss,speed_ms,0,blend_radius_m)
  movel([0.366879, -1.327364, -2.601345, -0.783680, 1.570796, 1.937675],accel_mss,speed_ms,0,blend_radius_m)
  movel([0.367180, -1.327824, -2.601053, -0.783512, 1.570796, 1.937976],accel_mss,speed_ms,0,blend_radius_m)
  movel([0.367684, -1.328091, -2.600884, -0.783414, 1.570796, 1.938480],accel_mss,speed_ms,0,blend_radius_m)
  movel([0.368319, -1.328150, -2.600846, -0.783393, 1.570796, 1.939115],accel_mss,speed_ms,0,blend_radius_m)
  movel([0.369026, -1.328056, -2.600906, -0.783427, 1.570796, 1.939822],accel_mss,speed_ms,0,blend_radius_m)
  movel([0.370518, -1.327557, -2.601222, -0.783609, 1.570796, 1.941314],accel_mss,speed_ms,0,blend_radius_m)
  movel([0.372420, -1.326616, -2.601819, -0.783954, 1.570796, 1.943216],accel_mss,speed_ms,0,blend_radius_m)
  movel([0.374257, -1.325428, -2.602569, -0.784391, 1.570796, 1.945053],accel_mss,speed_ms,0,blend_radius_m)
  movel([0.375978, -1.324034, -2.603448, -0.784907, 1.570796, 1.946774],accel_mss,speed_ms,0,blend_radius_m)
  movel([0.377529, -1.322469, -2.604432, -0.785488, 1.570796, 1.948326],accel_mss,speed_ms,0,blend_radius_m)
  movel([0.377980, -1.321898, -2.604790, -0.785701, 1.570796, 1.948776],accel_mss,speed_ms,0,blend_radius_m)
  movel([0.378215, -1.321320, -2.605151, -0.785917, 1.570796, 1.949011],accel_mss,speed_ms,0,blend_radius_m)
  movel([0.378135, -1.320914, -2.605405, -0.786069, 1.570796, 1.948931],accel_mss,speed_ms,0,blend_radius_m)
  movel([0.377887, -1.320608, -2.605597, -0.786184, 1.570796, 1.948683],accel_mss,speed_ms,0,blend_radius_m)
  movel([0.376822, -1.319803, -2.606100, -0.786487, 1.570796, 1.947618],accel_mss,speed_ms,0,blend_radius_m)
  movel([0.374629, -1.318541, -2.606886, -0.786963, 1.570796, 1.945425],accel_mss,speed_ms,0,blend_radius_m)
  movel([0.373735, -1.317564, -2.607493, -0.787332, 1.570796, 1.944532],accel_mss,speed_ms,0,blend_radius_m)
  movel([0.375862, -1.316051, -2.608430, -0.787907, 1.570796, 1.946659],accel_mss,speed_ms,0,blend_radius_m)
  movel([0.376980, -1.315466, -2.608792, -0.788131, 1.570796, 1.947776],accel_mss,speed_ms,0,blend_radius_m)
  movel([0.378104, -1.315058, -2.609045, -0.788287, 1.570796, 1.948900],accel_mss,speed_ms,0,blend_radius_m)
  movel([0.378856, -1.314916, -2.609132, -0.788341, 1.570796, 1.949653],accel_mss,speed_ms,0,blend_radius_m)
  movel([0.379619, -1.314884, -2.609152, -0.788353, 1.570796, 1.950415],accel_mss,speed_ms,0,blend_radius_m)
  movel([0.380928, -1.315127, -2.609002, -0.788260, 1.570796, 1.951724],accel_mss,speed_ms,0,blend_radius_m)
  movel([0.381539, -1.315644, -2.608682, -0.788063, 1.570796, 1.952335],accel_mss,speed_ms,0,blend_radius_m)
  movel([0.381668, -1.316031, -2.608443, -0.787915, 1.570796, 1.952464],accel_mss,speed_ms,0,blend_radius_m)
  movel([0.381635, -1.316492, -2.608158, -0.787739, 1.570796, 1.952431],accel_mss,speed_ms,0,blend_radius_m)
  movel([0.381346, -1.317129, -2.607763, -0.787497, 1.570796, 1.952142],accel_mss,speed_ms,0,blend_radius_m)
  movel([0.380854, -1.317730, -2.607390, -0.787269, 1.570796, 1.951650],accel_mss,speed_ms,0,blend_radius_m)
  movel([0.379565, -1.318775, -2.606740, -0.786874, 1.570796, 1.950361],accel_mss,speed_ms,0,blend_radius_m)
  speed_ms = 0.005
  movel([0.379565, -1.309823, -2.602454, -0.800112, 1.570796, 1.950361],accel_mss,speed_ms,0,blend_radius_m)
  speed_ms = 0.040
  movel([0.396456, -1.262957, -2.629851, -0.819581, 1.570796, 1.967252],accel_mss,speed_ms,0,blend_radius_m)
  speed_ms = 0.005
  movel([0.396456, -1.272161, -2.634347, -0.805881, 1.570796, 1.967252],accel_mss,speed_ms,0,blend_radius_m)
  speed_ms = 0.025
  movel([0.397325, -1.271763, -2.634571, -0.806055, 1.570796, 1.968121],accel_mss,speed_ms,0,blend_radius_m)
  movel([0.398176, -1.271516, -2.634709, -0.806163, 1.570796, 1.968972],accel_mss,speed_ms,0,blend_radius_m)
  movel([0.398993, -1.271412, -2.634768, -0.806209, 1.570796, 1.969789],accel_mss,speed_ms,0,blend_radius_m)
  movel([0.400468, -1.271599, -2.634663, -0.806127, 1.570796, 1.971265],accel_mss,speed_ms,0,blend_radius_m)
  movel([0.401097, -1.271872, -2.634509, -0.806008, 1.570796, 1.971893],accel_mss,speed_ms,0,blend_radius_m)
  movel([0.402060, -1.272730, -2.634026, -0.805632, 1.570796, 1.972857],accel_mss,speed_ms,0,blend_radius_m)
  movel([0.402608, -1.273911, -2.633360, -0.805118, 1.570796, 1.973405],accel_mss,speed_ms,0,blend_radius_m)
  movel([0.402816, -1.275301, -2.632574, -0.804514, 1.570796, 1.973612],accel_mss,speed_ms,0,blend_radius_m)
  movel([0.402748, -1.276830, -2.631706, -0.803853, 1.570796, 1.973544],accel_mss,speed_ms,0,blend_radius_m)
  movel([0.402471, -1.278427, -2.630796, -0.803165, 1.570796, 1.973267],accel_mss,speed_ms,0,blend_radius_m)
  movel([0.401764, -1.280899, -2.629382, -0.802108, 1.570796, 1.972560],accel_mss,speed_ms,0,blend_radius_m)
  movel([0.400753, -1.283400, -2.627944, -0.801045, 1.570796, 1.971550],accel_mss,speed_ms,0,blend_radius_m)
  movel([0.399458, -1.285891, -2.626503, -0.799995, 1.570796, 1.970255],accel_mss,speed_ms,0,blend_radius_m)
  movel([0.396374, -1.290632, -2.623740, -0.798017, 1.570796, 1.967171],accel_mss,speed_ms,0,blend_radius_m)
  movel([0.395862, -1.291755, -2.623081, -0.797553, 1.570796, 1.966658],accel_mss,speed_ms,0,blend_radius_m)
  movel([0.395718, -1.292802, -2.622465, -0.797122, 1.570796, 1.966514],accel_mss,speed_ms,0,blend_radius_m)
  movel([0.395972, -1.293573, -2.622011, -0.796805, 1.570796, 1.966768],accel_mss,speed_ms,0,blend_radius_m)
  movel([0.396450, -1.294199, -2.621641, -0.796548, 1.570796, 1.967246],accel_mss,speed_ms,0,blend_radius_m)
  movel([0.396975, -1.294800, -2.621286, -0.796302, 1.570796, 1.967771],accel_mss,speed_ms,0,blend_radius_m)
  movel([0.397363, -1.295494, -2.620876, -0.796019, 1.570796, 1.968159],accel_mss,speed_ms,0,blend_radius_m)
  movel([0.397477, -1.296253, -2.620426, -0.795710, 1.570796, 1.968273],accel_mss,speed_ms,0,blend_radius_m)
  movel([0.397384, -1.297101, -2.619923, -0.795365, 1.570796, 1.968180],accel_mss,speed_ms,0,blend_radius_m)
  movel([0.396839, -1.298907, -2.618847, -0.794634, 1.570796, 1.967635],accel_mss,speed_ms,0,blend_radius_m)
  movel([0.395796, -1.301518, -2.617286, -0.793585, 1.570796, 1.966593],accel_mss,speed_ms,0,blend_radius_m)
  movel([0.394602, -1.304123, -2.615719, -0.792547, 1.570796, 1.965398],accel_mss,speed_ms,0,blend_radius_m)
  movel([0.393256, -1.306710, -2.614154, -0.791525, 1.570796, 1.964052],accel_mss,speed_ms,0,blend_radius_m)
  movel([0.391770, -1.309274, -2.612594, -0.790521, 1.570796, 1.962566],accel_mss,speed_ms,0,blend_radius_m)
  movel([0.390148, -1.311800, -2.611049, -0.789540, 1.570796, 1.960945],accel_mss,speed_ms,0,blend_radius_m)
  movel([0.388402, -1.314281, -2.609524, -0.788584, 1.570796, 1.959199],accel_mss,speed_ms,0,blend_radius_m)
  movel([0.386532, -1.316707, -2.608024, -0.787658, 1.570796, 1.957328],accel_mss,speed_ms,0,blend_radius_m)
  movel([0.384547, -1.319072, -2.606555, -0.786762, 1.570796, 1.955344],accel_mss,speed_ms,0,blend_radius_m)
  movel([0.383210, -1.320514, -2.605655, -0.786219, 1.570796, 1.954007],accel_mss,speed_ms,0,blend_radius_m)
  movel([0.381746, -1.321849, -2.604820, -0.785720, 1.570796, 1.952543],accel_mss,speed_ms,0,blend_radius_m)
  movel([0.380183, -1.322928, -2.604144, -0.785318, 1.570796, 1.950980],accel_mss,speed_ms,0,blend_radius_m)
  movel([0.379375, -1.323320, -2.603897, -0.785172, 1.570796, 1.950172],accel_mss,speed_ms,0,blend_radius_m)
  movel([0.378551, -1.323595, -2.603724, -0.785069, 1.570796, 1.949348],accel_mss,speed_ms,0,blend_radius_m)
  speed_ms = 0.005
  movel([0.378551, -1.314671, -2.599460, -0.798258, 1.570796, 1.949348],accel_mss,speed_ms,0,blend_radius_m)
  speed_ms = 0.040
  movel([0.373988, -1.318367, -2.597157, -0.796865, 1.570796, 1.944785],accel_mss,speed_ms,0,blend_radius_m)
  speed_ms = 0.005
  movel([0.373988, -1.327269, -2.601405, -0.783715, 1.570796, 1.944785],accel_mss,speed_ms,0,blend_radius_m)
  speed_ms = 0.025
  movel([0.374067, -1.327774, -2.601085, -0.783530, 1.570796, 1.944863],accel_mss,speed_ms,0,blend_radius_m)
  movel([0.373867, -1.328373, -2.600705, -0.783311, 1.570796, 1.944663],accel_mss,speed_ms,0,blend_radius_m)
  movel([0.373459, -1.328983, -2.600317, -0.783089, 1.570796, 1.944256],accel_mss,speed_ms,0,blend_radius_m)
  movel([0.372910, -1.329520, -2.599975, -0.782894, 1.570796, 1.943706],accel_mss,speed_ms,0,blend_radius_m)
  movel([0.372159, -1.329965, -2.599691, -0.782732, 1.570796, 1.942956],accel_mss,speed_ms,0,blend_radius_m)
  movel([0.371404, -1.330237, -2.599518, -0.782634, 1.570796, 1.942200],accel_mss,speed_ms,0,blend_radius_m)
  movel([0.370665, -1.330476, -2.599366, -0.782547, 1.570796, 1.941462],accel_mss,speed_ms,0,blend_radius_m)
  movel([0.369977, -1.330830, -2.599140, -0.782419, 1.570796, 1.940773],accel_mss,speed_ms,0,blend_radius_m)
  movel([0.369216, -1.331639, -2.598623, -0.782127, 1.570796, 1.940013],accel_mss,speed_ms,0,blend_radius_m)
  movel([0.368860, -1.332082, -2.598340, -0.781968, 1.570796, 1.939657],accel_mss,speed_ms,0,blend_radius_m)
  movel([0.368392, -1.332504, -2.598069, -0.781816, 1.570796, 1.939188],accel_mss,speed_ms,0,blend_radius_m)
  movel([0.366956, -1.333415, -2.597485, -0.781489, 1.570796, 1.937753],accel_mss,speed_ms,0,blend_radius_m)
  movel([0.365524, -1.334099, -2.597045, -0.781245, 1.570796, 1.936320],accel_mss,speed_ms,0,blend_radius_m)
  movel([0.364083, -1.334585, -2.596732, -0.781071, 1.570796, 1.934879],accel_mss,speed_ms,0,blend_radius_m)
  movel([0.362620, -1.334913, -2.596521, -0.780954, 1.570796, 1.933416],accel_mss,speed_ms,0,blend_radius_m)
  movel([0.363390, -1.334667, -2.596680, -0.781042, 1.570796, 1.934186],accel_mss,speed_ms,0,blend_radius_m)
  movel([0.364136, -1.334534, -2.596765, -0.781089, 1.570796, 1.934932],accel_mss,speed_ms,0,blend_radius_m)
  movel([0.364781, -1.334639, -2.596698, -0.781052, 1.570796, 1.935577],accel_mss,speed_ms,0,blend_radius_m)
  movel([0.365146, -1.335050, -2.596433, -0.780906, 1.570796, 1.935942],accel_mss,speed_ms,0,blend_radius_m)
  movel([0.365074, -1.335695, -2.596018, -0.780677, 1.570796, 1.935870],accel_mss,speed_ms,0,blend_radius_m)
  movel([0.364665, -1.336380, -2.595575, -0.780434, 1.570796, 1.935461],accel_mss,speed_ms,0,blend_radius_m)
  movel([0.364051, -1.336973, -2.595192, -0.780224, 1.570796, 1.934848],accel_mss,speed_ms,0,blend_radius_m)
  movel([0.362189, -1.338184, -2.594407, -0.779797, 1.570796, 1.932986],accel_mss,speed_ms,0,blend_radius_m)
  movel([0.360995, -1.338773, -2.594025, -0.779591, 1.570796, 1.931792],accel_mss,speed_ms,0,blend_radius_m)
  movel([0.359796, -1.339236, -2.593725, -0.779429, 1.570796, 1.930592],accel_mss,speed_ms,0,blend_radius_m)
  movel([0.358603, -1.339564, -2.593511, -0.779314, 1.570796, 1.929399],accel_mss,speed_ms,0,blend_radius_m)
  movel([0.359929, -1.339375, -2.593634, -0.779380, 1.570796, 1.930726],accel_mss,speed_ms,0,blend_radius_m)
  movel([0.361336, -1.339014, -2.593869, -0.779506, 1.570796, 1.932132],accel_mss,speed_ms,0,blend_radius_m)
  movel([0.362708, -1.338690, -2.594079, -0.779620, 1.570796, 1.933504],accel_mss,speed_ms,0,blend_radius_m)
  movel([0.363934, -1.338599, -2.594139, -0.779652, 1.570796, 1.934730],accel_mss,speed_ms,0,blend_radius_m)
  movel([0.364250, -1.338727, -2.594055, -0.779607, 1.570796, 1.935047],accel_mss,speed_ms,0,blend_radius_m)
  movel([0.364221, -1.338988, -2.593886, -0.779515, 1.570796, 1.935017],accel_mss,speed_ms,0,blend_radius_m)
  movel([0.363382, -1.340043, -2.593199, -0.779146, 1.570796, 1.934179],accel_mss,speed_ms,0,blend_radius_m)
  movel([0.362643, -1.340745, -2.592742, -0.778902, 1.570796, 1.933439],accel_mss,speed_ms,0,blend_radius_m)
  movel([0.361836, -1.341371, -2.592334, -0.778684, 1.570796, 1.932632],accel_mss,speed_ms,0,blend_radius_m)
  movel([0.360982, -1.341903, -2.591987, -0.778500, 1.570796, 1.931778],accel_mss,speed_ms,0,blend_radius_m)
  movel([0.361400, -1.341739, -2.592093, -0.778556, 1.570796, 1.932197],accel_mss,speed_ms,0,blend_radius_m)
  movel([0.361850, -1.341682, -2.592131, -0.778576, 1.570796, 1.932646],accel_mss,speed_ms,0,blend_radius_m)
  movel([0.362789, -1.341835, -2.592031, -0.778523, 1.570796, 1.933585],accel_mss,speed_ms,0,blend_radius_m)
  movel([0.363680, -1.342269, -2.591747, -0.778373, 1.570796, 1.934477],accel_mss,speed_ms,0,blend_radius_m)
  movel([0.364415, -1.342889, -2.591341, -0.778158, 1.570796, 1.935212],accel_mss,speed_ms,0,blend_radius_m)
  movel([0.364885, -1.343601, -2.590874, -0.777913, 1.570796, 1.935681],accel_mss,speed_ms,0,blend_radius_m)
  movel([0.364980, -1.344308, -2.590411, -0.777670, 1.570796, 1.935776],accel_mss,speed_ms,0,blend_radius_m)
  movel([0.364853, -1.344629, -2.590200, -0.777560, 1.570796, 1.935649],accel_mss,speed_ms,0,blend_radius_m)
  movel([0.364591, -1.344912, -2.590014, -0.777463, 1.570796, 1.935387],accel_mss,speed_ms,0,blend_radius_m)
  movel([0.364182, -1.345149, -2.589858, -0.777382, 1.570796, 1.934978],accel_mss,speed_ms,0,blend_radius_m)
  movel([0.363610, -1.345325, -2.589742, -0.777322, 1.570796, 1.934406],accel_mss,speed_ms,0,blend_radius_m)
  movel([0.363000, -1.345353, -2.589724, -0.777312, 1.570796, 1.933796],accel_mss,speed_ms,0,blend_radius_m)
  movel([0.360836, -1.344651, -2.590185, -0.777553, 1.570796, 1.931632],accel_mss,speed_ms,0,blend_radius_m)
  movel([0.359985, -1.344431, -2.590330, -0.777628, 1.570796, 1.930781],accel_mss,speed_ms,0,blend_radius_m)
  movel([0.359045, -1.344374, -2.590368, -0.777648, 1.570796, 1.929841],accel_mss,speed_ms,0,blend_radius_m)
  movel([0.357337, -1.344694, -2.590157, -0.777538, 1.570796, 1.928133],accel_mss,speed_ms,0,blend_radius_m)
  movel([0.355594, -1.345133, -2.589869, -0.777388, 1.570796, 1.926391],accel_mss,speed_ms,0,blend_radius_m)
  movel([0.354745, -1.345213, -2.589816, -0.777360, 1.570796, 1.925542],accel_mss,speed_ms,0,blend_radius_m)
  movel([0.353980, -1.345115, -2.589880, -0.777394, 1.570796, 1.924776],accel_mss,speed_ms,0,blend_radius_m)
  movel([0.353402, -1.344805, -2.590084, -0.777500, 1.570796, 1.924198],accel_mss,speed_ms,0,blend_radius_m)
  movel([0.353111, -1.344250, -2.590449, -0.777690, 1.570796, 1.923907],accel_mss,speed_ms,0,blend_radius_m)
  movel([0.354048, -1.343478, -2.590955, -0.777955, 1.570796, 1.924844],accel_mss,speed_ms,0,blend_radius_m)
  movel([0.355043, -1.342795, -2.591403, -0.778191, 1.570796, 1.925839],accel_mss,speed_ms,0,blend_radius_m)
  speed_ms = 0.005
  movel([0.355043, -1.333988, -2.587223, -0.791177, 1.570796, 1.925839],accel_mss,speed_ms,0,blend_radius_m)
  speed_ms = 0.040
  movel([0.361691, -1.341694, -2.582203, -0.788492, 1.570796, 1.932487],accel_mss,speed_ms,0,blend_radius_m)
  speed_ms = 0.005
  movel([0.361691, -1.350453, -2.586349, -0.775587, 1.570796, 1.932487],accel_mss,speed_ms,0,blend_radius_m)
  speed_ms = 0.025
  movel([0.362348, -1.349898, -2.586718, -0.775773, 1.570796, 1.933144],accel_mss,speed_ms,0,blend_radius_m)
  movel([0.363111, -1.349601, -2.586915, -0.775873, 1.570796, 1.933908],accel_mss,speed_ms,0,blend_radius_m)
  movel([0.363859, -1.349559, -2.586943, -0.775887, 1.570796, 1.934656],accel_mss,speed_ms,0,blend_radius_m)
  movel([0.364464, -1.349770, -2.586803, -0.775816, 1.570796, 1.935260],accel_mss,speed_ms,0,blend_radius_m)
  movel([0.364865, -1.350180, -2.586530, -0.775679, 1.570796, 1.935662],accel_mss,speed_ms,0,blend_radius_m)
  movel([0.365116, -1.350709, -2.586178, -0.775502, 1.570796, 1.935912],accel_mss,speed_ms,0,blend_radius_m)
  movel([0.365357, -1.351940, -2.585358, -0.775091, 1.570796, 1.936153],accel_mss,speed_ms,0,blend_radius_m)
  movel([0.365972, -1.351175, -2.585868, -0.775346, 1.570796, 1.936768],accel_mss,speed_ms,0,blend_radius_m)
  movel([0.366388, -1.350358, -2.586412, -0.775619, 1.570796, 1.937185],accel_mss,speed_ms,0,blend_radius_m)
  movel([0.366573, -1.349560, -2.586942, -0.775887, 1.570796, 1.937369],accel_mss,speed_ms,0,blend_radius_m)
  movel([0.366505, -1.348842, -2.587418, -0.776128, 1.570796, 1.937301],accel_mss,speed_ms,0,blend_radius_m)
  movel([0.366873, -1.349210, -2.587174, -0.776005, 1.570796, 1.937669],accel_mss,speed_ms,0,blend_radius_m)
  movel([0.367116, -1.349666, -2.586872, -0.775851, 1.570796, 1.937912],accel_mss,speed_ms,0,blend_radius_m)
  movel([0.367295, -1.350774, -2.586135, -0.775480, 1.570796, 1.938091],accel_mss,speed_ms,0,blend_radius_m)
  movel([0.367188, -1.352042, -2.585290, -0.775057, 1.570796, 1.937984],accel_mss,speed_ms,0,blend_radius_m)
  movel([0.366924, -1.353353, -2.584414, -0.774623, 1.570796, 1.937720],accel_mss,speed_ms,0,blend_radius_m)
  movel([0.366429, -1.354796, -2.583446, -0.774147, 1.570796, 1.937226],accel_mss,speed_ms,0,blend_radius_m)
  movel([0.365752, -1.356154, -2.582533, -0.773702, 1.570796, 1.936548],accel_mss,speed_ms,0,blend_radius_m)
  movel([0.365054, -1.357483, -2.581638, -0.773269, 1.570796, 1.935850],accel_mss,speed_ms,0,blend_radius_m)
  movel([0.364495, -1.358842, -2.580719, -0.772828, 1.570796, 1.935291],accel_mss,speed_ms,0,blend_radius_m)
  movel([0.364072, -1.357929, -2.581336, -0.773124, 1.570796, 1.934868],accel_mss,speed_ms,0,blend_radius_m)
  movel([0.363392, -1.357221, -2.581814, -0.773354, 1.570796, 1.934188],accel_mss,speed_ms,0,blend_radius_m)
  movel([0.362472, -1.356759, -2.582126, -0.773504, 1.570796, 1.933268],accel_mss,speed_ms,0,blend_radius_m)
  movel([0.361324, -1.356584, -2.582244, -0.773561, 1.570796, 1.932120],accel_mss,speed_ms,0,blend_radius_m)
  speed_ms = 0.005
  movel([0.361324, -1.347864, -2.578126, -0.786399, 1.570796, 1.932120],accel_mss,speed_ms,0,blend_radius_m)
  speed_ms = 0.040
  movel([0.361828, -1.352455, -2.575058, -0.784876, 1.570796, 1.932624],accel_mss,speed_ms,0,blend_radius_m)
  speed_ms = 0.005
  movel([0.361828, -1.361145, -2.579156, -0.772088, 1.570796, 1.932624],accel_mss,speed_ms,0,blend_radius_m)
  speed_ms = 0.025
  movel([0.361728, -1.362939, -2.577934, -0.771516, 1.570796, 1.932524],accel_mss,speed_ms,0,blend_radius_m)
  movel([0.361919, -1.364612, -2.576790, -0.770987, 1.570796, 1.932715],accel_mss,speed_ms,0,blend_radius_m)
  movel([0.362508, -1.366020, -2.575824, -0.770545, 1.570796, 1.933305],accel_mss,speed_ms,0,blend_radius_m)
  movel([0.362989, -1.366579, -2.575439, -0.770370, 1.570796, 1.933785],accel_mss,speed_ms,0,blend_radius_m)
  movel([0.363612, -1.367021, -2.575136, -0.770233, 1.570796, 1.934409],accel_mss,speed_ms,0,blend_radius_m)
  movel([0.364670, -1.367391, -2.574881, -0.770117, 1.570796, 1.935466],accel_mss,speed_ms,0,blend_radius_m)
  movel([0.365870, -1.367503, -2.574804, -0.770082, 1.570796, 1.936666],accel_mss,speed_ms,0,blend_radius_m)
  movel([0.367181, -1.367419, -2.574861, -0.770109, 1.570796, 1.937978],accel_mss,speed_ms,0,blend_radius_m)
  movel([0.368573, -1.367199, -2.575013, -0.770177, 1.570796, 1.939369],accel_mss,speed_ms,0,blend_radius_m)
  movel([0.371467, -1.366585, -2.575435, -0.770368, 1.570796, 1.942264],accel_mss,speed_ms,0,blend_radius_m)
  movel([0.374296, -1.366145, -2.575738, -0.770506, 1.570796, 1.945092],accel_mss,speed_ms,0,blend_radius_m)
  movel([0.375819, -1.366154, -2.575732, -0.770503, 1.570796, 1.946615],accel_mss,speed_ms,0,blend_radius_m)
  movel([0.377217, -1.366397, -2.575565, -0.770427, 1.570796, 1.948013],accel_mss,speed_ms,0,blend_radius_m)
  movel([0.378467, -1.366858, -2.575248, -0.770283, 1.570796, 1.949264],accel_mss,speed_ms,0,blend_radius_m)
  movel([0.379548, -1.367523, -2.574790, -0.770076, 1.570796, 1.950344],accel_mss,speed_ms,0,blend_radius_m)
  movel([0.380440, -1.368370, -2.574206, -0.769813, 1.570796, 1.951237],accel_mss,speed_ms,0,blend_radius_m)
  movel([0.381123, -1.369387, -2.573503, -0.769499, 1.570796, 1.951919],accel_mss,speed_ms,0,blend_radius_m)
  movel([0.381572, -1.370554, -2.572695, -0.769140, 1.570796, 1.952369],accel_mss,speed_ms,0,blend_radius_m)
  movel([0.381775, -1.371852, -2.571794, -0.768744, 1.570796, 1.952571],accel_mss,speed_ms,0,blend_radius_m)
  speed_ms = 0.005
  movel([0.381775, -1.363232, -2.567742, -0.781414, 1.570796, 1.952571],accel_mss,speed_ms,0,blend_radius_m)
  speed_ms = 0.040
  movel([0.359238, -1.338381, -2.584371, -0.789636, 1.570796, 1.930034],accel_mss,speed_ms,0,blend_radius_m)
  speed_ms = 0.005
  movel([0.359238, -1.347161, -2.588531, -0.776697, 1.570796, 1.930034],accel_mss,speed_ms,0,blend_radius_m)
  speed_ms = 0.025
  movel([0.359845, -1.347603, -2.588239, -0.776547, 1.570796, 1.930641],accel_mss,speed_ms,0,blend_radius_m)
  movel([0.360242, -1.348213, -2.587836, -0.776341, 1.570796, 1.931038],accel_mss,speed_ms,0,blend_radius_m)
  movel([0.360277, -1.348619, -2.587566, -0.776203, 1.570796, 1.931074],accel_mss,speed_ms,0,blend_radius_m)
  movel([0.360167, -1.349072, -2.587266, -0.776051, 1.570796, 1.930964],accel_mss,speed_ms,0,blend_radius_m)
  movel([0.359916, -1.349517, -2.586971, -0.775901, 1.570796, 1.930712],accel_mss,speed_ms,0,blend_radius_m)
  movel([0.359523, -1.349899, -2.586717, -0.775773, 1.570796, 1.930319],accel_mss,speed_ms,0,blend_radius_m)
  movel([0.358663, -1.350431, -2.586363, -0.775595, 1.570796, 1.929459],accel_mss,speed_ms,0,blend_radius_m)
  movel([0.358328, -1.350811, -2.586110, -0.775468, 1.570796, 1.929124],accel_mss,speed_ms,0,blend_radius_m)
  movel([0.358144, -1.351235, -2.585828, -0.775326, 1.570796, 1.928941],accel_mss,speed_ms,0,blend_radius_m)
  movel([0.358112, -1.352066, -2.585273, -0.775049, 1.570796, 1.928908],accel_mss,speed_ms,0,blend_radius_m)
  movel([0.358346, -1.352917, -2.584705, -0.774767, 1.570796, 1.929142],accel_mss,speed_ms,0,blend_radius_m)
  movel([0.358741, -1.353665, -2.584205, -0.774519, 1.570796, 1.929537],accel_mss,speed_ms,0,blend_radius_m)
  movel([0.359287, -1.354302, -2.583778, -0.774309, 1.570796, 1.930083],accel_mss,speed_ms,0,blend_radius_m)
  movel([0.359971, -1.354808, -2.583438, -0.774143, 1.570796, 1.930767],accel_mss,speed_ms,0,blend_radius_m)
  movel([0.359211, -1.355657, -2.582868, -0.773864, 1.570796, 1.930007],accel_mss,speed_ms,0,blend_radius_m)
  movel([0.358601, -1.356547, -2.582269, -0.773573, 1.570796, 1.929397],accel_mss,speed_ms,0,blend_radius_m)
  movel([0.358123, -1.357466, -2.581649, -0.773274, 1.570796, 1.928920],accel_mss,speed_ms,0,blend_radius_m)
  movel([0.357762, -1.358402, -2.581017, -0.772970, 1.570796, 1.928558],accel_mss,speed_ms,0,blend_radius_m)
  movel([0.357327, -1.360277, -2.579746, -0.772366, 1.570796, 1.928123],accel_mss,speed_ms,0,blend_radius_m)
  movel([0.357176, -1.362080, -2.578519, -0.771789, 1.570796, 1.927973],accel_mss,speed_ms,0,blend_radius_m)
  movel([0.357067, -1.363810, -2.577338, -0.771240, 1.570796, 1.927863],accel_mss,speed_ms,0,blend_radius_m)
  movel([0.356873, -1.364698, -2.576731, -0.770960, 1.570796, 1.927670],accel_mss,speed_ms,0,blend_radius_m)
  movel([0.356501, -1.365601, -2.576111, -0.770676, 1.570796, 1.927298],accel_mss,speed_ms,0,blend_radius_m)
  movel([0.355871, -1.366494, -2.575498, -0.770397, 1.570796, 1.926667],accel_mss,speed_ms,0,blend_radius_m)
  movel([0.355024, -1.367265, -2.574968, -0.770156, 1.570796, 1.925820],accel_mss,speed_ms,0,blend_radius_m)
  movel([0.354078, -1.367787, -2.574608, -0.769994, 1.570796, 1.924875],accel_mss,speed_ms,0,blend_radius_m)
  movel([0.353157, -1.367928, -2.574511, -0.769950, 1.570796, 1.923953],accel_mss,speed_ms,0,blend_radius_m)
  movel([0.353394, -1.368637, -2.574021, -0.769731, 1.570796, 1.924191],accel_mss,speed_ms,0,blend_radius_m)
  movel([0.353487, -1.370236, -2.572915, -0.769238, 1.570796, 1.924283],accel_mss,speed_ms,0,blend_radius_m)
  movel([0.353346, -1.371098, -2.572318, -0.768974, 1.570796, 1.924143],accel_mss,speed_ms,0,blend_radius_m)
  movel([0.352717, -1.372872, -2.571084, -0.768433, 1.570796, 1.923513],accel_mss,speed_ms,0,blend_radius_m)
  movel([0.352233, -1.373755, -2.570468, -0.768166, 1.570796, 1.923030],accel_mss,speed_ms,0,blend_radius_m)
  movel([0.351639, -1.374619, -2.569864, -0.767905, 1.570796, 1.922436],accel_mss,speed_ms,0,blend_radius_m)
  speed_ms = 0.005
  movel([0.351639, -1.366019, -2.565825, -0.780546, 1.570796, 1.922436],accel_mss,speed_ms,0,blend_radius_m)
  speed_ms = 0.040
  movel([0.347238, -1.365916, -2.565895, -0.780577, 1.570796, 1.918034],accel_mss,speed_ms,0,blend_radius_m)
  speed_ms = 0.005
  movel([0.347238, -1.374518, -2.569935, -0.767936, 1.570796, 1.918034],accel_mss,speed_ms,0,blend_radius_m)
  speed_ms = 0.025
  movel([0.348190, -1.382732, -2.564146, -0.765511, 1.570796, 1.918986],accel_mss,speed_ms,0,blend_radius_m)
  movel([0.348182, -1.383778, -2.563401, -0.765209, 1.570796, 1.918978],accel_mss,speed_ms,0,blend_radius_m)
  movel([0.348003, -1.384315, -2.563019, -0.765055, 1.570796, 1.918799],accel_mss,speed_ms,0,blend_radius_m)
  movel([0.347631, -1.384822, -2.562657, -0.764910, 1.570796, 1.918427],accel_mss,speed_ms,0,blend_radius_m)
  movel([0.346522, -1.385757, -2.561989, -0.764643, 1.570796, 1.917319],accel_mss,speed_ms,0,blend_radius_m)
  movel([0.346243, -1.386337, -2.561574, -0.764478, 1.570796, 1.917039],accel_mss,speed_ms,0,blend_radius_m)
  movel([0.346216, -1.386900, -2.561171, -0.764318, 1.570796, 1.917013],accel_mss,speed_ms,0,blend_radius_m)
  movel([0.346487, -1.387707, -2.560592, -0.764090, 1.570796, 1.917284],accel_mss,speed_ms,0,blend_radius_m)
  movel([0.347023, -1.388384, -2.560106, -0.763899, 1.570796, 1.917819],accel_mss,speed_ms,0,blend_radius_m)
  movel([0.348262, -1.389564, -2.559257, -0.763568, 1.570796, 1.919058],accel_mss,speed_ms,0,blend_radius_m)
  movel([0.348868, -1.390503, -2.558579, -0.763306, 1.570796, 1.919664],accel_mss,speed_ms,0,blend_radius_m)
  movel([0.349474, -1.391987, -2.557507, -0.762895, 1.570796, 1.920271],accel_mss,speed_ms,0,blend_radius_m)
  movel([0.349582, -1.392730, -2.556968, -0.762691, 1.570796, 1.920379],accel_mss,speed_ms,0,blend_radius_m)
  movel([0.349464, -1.393364, -2.556508, -0.762517, 1.570796, 1.920260],accel_mss,speed_ms,0,blend_radius_m)
  movel([0.349294, -1.393615, -2.556326, -0.762448, 1.570796, 1.920090],accel_mss,speed_ms,0,blend_radius_m)
  movel([0.349038, -1.393806, -2.556187, -0.762396, 1.570796, 1.919834],accel_mss,speed_ms,0,blend_radius_m)
  movel([0.348227, -1.393980, -2.556061, -0.762348, 1.570796, 1.919023],accel_mss,speed_ms,0,blend_radius_m)
  movel([0.348190, -1.394646, -2.555576, -0.762167, 1.570796, 1.918986],accel_mss,speed_ms,0,blend_radius_m)
  movel([0.348361, -1.395335, -2.555075, -0.761980, 1.570796, 1.919157],accel_mss,speed_ms,0,blend_radius_m)
  movel([0.349135, -1.396694, -2.554082, -0.761612, 1.570796, 1.919931],accel_mss,speed_ms,0,blend_radius_m)
  movel([0.351071, -1.398815, -2.552529, -0.761045, 1.570796, 1.921867],accel_mss,speed_ms,0,blend_radius_m)
  movel([0.352265, -1.399665, -2.551905, -0.760819, 1.570796, 1.923061],accel_mss,speed_ms,0,blend_radius_m)
  movel([0.353639, -1.400431, -2.551342, -0.760617, 1.570796, 1.924436],accel_mss,speed_ms,0,blend_radius_m)
  movel([0.354826, -1.401333, -2.550676, -0.760380, 1.570796, 1.925622],accel_mss,speed_ms,0,blend_radius_m)
  movel([0.355234, -1.401903, -2.550256, -0.760230, 1.570796, 1.926031],accel_mss,speed_ms,0,blend_radius_m)
  movel([0.355458, -1.402588, -2.549750, -0.760051, 1.570796, 1.926255],accel_mss,speed_ms,0,blend_radius_m)
  movel([0.355448, -1.402997, -2.549447, -0.759945, 1.570796, 1.926244],accel_mss,speed_ms,0,blend_radius_m)
  movel([0.355305, -1.403430, -2.549126, -0.759832, 1.570796, 1.926101],accel_mss,speed_ms,0,blend_radius_m)
  movel([0.355033, -1.403803, -2.548850, -0.759736, 1.570796, 1.925829],accel_mss,speed_ms,0,blend_radius_m)
  movel([0.354631, -1.404024, -2.548686, -0.759679, 1.570796, 1.925428],accel_mss,speed_ms,0,blend_radius_m)
  movel([0.354024, -1.403933, -2.548754, -0.759702, 1.570796, 1.924820],accel_mss,speed_ms,0,blend_radius_m)
  movel([0.351655, -1.402668, -2.549691, -0.760031, 1.570796, 1.922451],accel_mss,speed_ms,0,blend_radius_m)
  movel([0.349595, -1.401079, -2.550864, -0.760446, 1.570796, 1.920391],accel_mss,speed_ms,0,blend_radius_m)
  movel([0.349319, -1.401514, -2.550543, -0.760332, 1.570796, 1.920115],accel_mss,speed_ms,0,blend_radius_m)
  movel([0.349162, -1.401955, -2.550217, -0.760217, 1.570796, 1.919958],accel_mss,speed_ms,0,blend_radius_m)
  movel([0.349160, -1.402846, -2.549559, -0.759984, 1.570796, 1.919956],accel_mss,speed_ms,0,blend_radius_m)
  movel([0.349492, -1.403721, -2.548911, -0.759757, 1.570796, 1.920288],accel_mss,speed_ms,0,blend_radius_m)
  movel([0.350058, -1.404564, -2.548286, -0.759540, 1.570796, 1.920854],accel_mss,speed_ms,0,blend_radius_m)
  movel([0.351526, -1.406039, -2.547189, -0.759161, 1.570796, 1.922323],accel_mss,speed_ms,0,blend_radius_m)
  movel([0.352807, -1.407079, -2.546414, -0.758896, 1.570796, 1.923603],accel_mss,speed_ms,0,blend_radius_m)
  movel([0.353218, -1.407518, -2.546086, -0.758785, 1.570796, 1.924014],accel_mss,speed_ms,0,blend_radius_m)
  movel([0.353302, -1.407798, -2.545877, -0.758714, 1.570796, 1.924098],accel_mss,speed_ms,0,blend_radius_m)
  movel([0.353235, -1.408127, -2.545631, -0.758631, 1.570796, 1.924031],accel_mss,speed_ms,0,blend_radius_m)
  movel([0.353004, -1.408478, -2.545368, -0.758542, 1.570796, 1.923800],accel_mss,speed_ms,0,blend_radius_m)
  movel([0.352724, -1.408689, -2.545211, -0.758489, 1.570796, 1.923521],accel_mss,speed_ms,0,blend_radius_m)
  movel([0.352084, -1.408836, -2.545101, -0.758452, 1.570796, 1.922880],accel_mss,speed_ms,0,blend_radius_m)
  movel([0.351196, -1.408954, -2.545012, -0.758422, 1.570796, 1.921992],accel_mss,speed_ms,0,blend_radius_m)
  movel([0.350992, -1.409119, -2.544889, -0.758381, 1.570796, 1.921789],accel_mss,speed_ms,0,blend_radius_m)
  movel([0.350845, -1.409427, -2.544658, -0.758304, 1.570796, 1.921641],accel_mss,speed_ms,0,blend_radius_m)
  movel([0.350832, -1.409758, -2.544410, -0.758221, 1.570796, 1.921628],accel_mss,speed_ms,0,blend_radius_m)
  movel([0.351090, -1.410430, -2.543906, -0.758053, 1.570796, 1.921887],accel_mss,speed_ms,0,blend_radius_m)
  movel([0.351887, -1.411506, -2.543097, -0.757786, 1.570796, 1.922683],accel_mss,speed_ms,0,blend_radius_m)
  movel([0.355713, -1.415710, -2.539920, -0.756759, 1.570796, 1.926510],accel_mss,speed_ms,0,blend_radius_m)
  movel([0.356016, -1.416194, -2.539552, -0.756642, 1.570796, 1.926812],accel_mss,speed_ms,0,blend_radius_m)
  movel([0.356172, -1.416763, -2.539120, -0.756506, 1.570796, 1.926968],accel_mss,speed_ms,0,blend_radius_m)
  movel([0.356086, -1.417358, -2.538667, -0.756363, 1.570796, 1.926882],accel_mss,speed_ms,0,blend_radius_m)
  movel([0.355659, -1.417922, -2.538238, -0.756229, 1.570796, 1.926455],accel_mss,speed_ms,0,blend_radius_m)
  movel([0.355048, -1.418250, -2.537988, -0.756151, 1.570796, 1.925844],accel_mss,speed_ms,0,blend_radius_m)
  movel([0.354427, -1.418298, -2.537951, -0.756140, 1.570796, 1.925223],accel_mss,speed_ms,0,blend_radius_m)
  movel([0.353842, -1.418150, -2.538064, -0.756175, 1.570796, 1.924638],accel_mss,speed_ms,0,blend_radius_m)
